Omron Sysmac Studio project Battery_System_Before_Test (Sysmac Studio 1.53.0.9, StandardProject)

# Controller new_Controller_0: NX102-1020 version 1.33
Units and slaves: 노드1 : NX-ECC203 (E005); 유니트 1 : NX-ID6142-6 (N8); 유니트 2 : NX-OD6121-6 (N9); 유니트 1 : NX-PF0730 (N1); 유니트 2 : NX-ILM400 (N2); 유니트 4 : NX-SID800 (N10); 유니트 5 : NX-SOD400 (N11)
Task PrimaryTask (priority 4, period or condition 2000): Program0, SlotTableProc

TYPE Slot_info : STRUCT
    SOC : UINT;  (* 배터리 잔량 % *)
    Status : INT;  (* 0 = 비어 있음 / 1 = 충전 중 / 2 = 불량 *)
    IO : WORD;  (* 로봇 신호 *)
END_STRUCT END_TYPE
TYPE U_IO16 : UNION
    W : WORD;
    B : ARRAY[0..15] OF BOOL;
END_UNION END_TYPE
TYPE S_RobotIO : STRUCT
    IO : U_IO16;
END_STRUCT END_TYPE

VAR_GLOBAL RETAIN
    Slot_No : ARRAY[1..6] OF Slot_Info := [(SOC := 16#0, Status := 1, IO := 16#01), (SOC := 16#0, Status := 1, IO := 16#02), (SOC := 16#0, Status := 1, IO := 16#04), (SOC := 16#0, Status := 1, IO := 16#08), (SOC := 16#0, Status := 1, IO := 16#10), (SOC := 16#0, Status := 1, IO := 16#20)];
END_VAR
VAR_GLOBAL
    Vision_Trigger : BOOL;  (* at ECAT://node#4/Line0 Trigger *)
    Vision_BC_Data : DINT;  (* at ECAT://node#4/Line0 DINT Result Data 0 *)
    Vision_Counter : DINT;  (* at ECAT://node#4/Line0 DINT Result Data 1 *)
    Robot_Send : S_RobotIO;
    Robot_Recv : S_RobotIO;
    MFC_HR : ARRAY[0..99] OF WORD;  (* PLC > MFC *)
    Arduino_HR : ARRAY[0..99] OF WORD;  (* Arduino > PLC *)
    Robot_In : ARRAY[0..237] OF WORD;  (* Robot > PLC; network input *)
    Robot_Out : ARRAY[0..105] OF WORD;  (* PLC > Robot; network output *)
    E_RST : BOOL;  (* Error Reset *)
    H_Rent_PB : BOOL;
    H_Card_Can_PB : BOOL;
    H_LowBatt_OK_PB : BOOL;
    H_LowBatt_Can_PB : BOOL;
    STP_D_SS : BOOL;  (* at ECAT://node#[1,1]/Input Bit 32 bits/Input Bit 16 *)
    STP_U_SS : BOOL;  (* at ECAT://node#[1,1]/Input Bit 32 bits/Input Bit 15 *)
    Detect_Home_SS : BOOL;  (* at ECAT://node#[1,1]/Input Bit 32 bits/Input Bit 22 *)
    Detect_STP_SS : BOOL;  (* at ECAT://node#[1,1]/Input Bit 32 bits/Input Bit 21 *)
    H_Vis_Rty_PB : BOOL;
    H_Vis_Home_PB : BOOL;
    H_Rtn_PB : BOOL;
    H_Rtn_Can_PB : BOOL;
    H_Refund_Can_PB : BOOL;
    H_Pop_Card : BOOL;
    H_pop_Wait_Rent : BOOL;
    H_Pop_LowBatt : BOOL;
    H_Pop_ContAdmin : BOOL;
    H_Pop_Rent_Done : BOOL;
    H_Pop_Place_Batt : BOOL;
    H_Pop_ReplBatt : BOOL;
    H_Pop_Refund : BOOL;
    H_Pop_RtnDone : BOOL;
    H_Pop_Equip_Running : BOOL;
    STP_SOL : BOOL;  (* at ECAT://node#[1,2]/Output Bit 32 bits/Output Bit 11 *)
    H_Scr_Main : BOOL;
    MotS_Status : WORD;  (* at ECAT://node#2/Status *)
    MotS : WORD;  (* at ECAT://node#2/Command *)
    MotM : WORD;  (* at ECAT://node#3/Command *)
    MotM_Status : WORD;  (* at ECAT://node#3/Status *)
    Batt_UseTime : ARRAY[1..6] OF TIME;
    Batt_Max_SOC : UINT;
    H_Pop_PayFail : BOOL;
    H_PayRty_PB : BOOL;
    H_PayFail_Home_PB : BOOL;
    Rtn_BC_IDX : DINT;
    Batt_Refund : LINT;
    H_Rst_PB : BOOL;
    H_Admin_PB : BOOL;
    H_Pop_Admin : BOOL;
    H_Admin_Home_PB : BOOL;
    RobotDone : BOOL;  (* 로봇 작업 완료 *)
    RobotMode : INT;  (* 1 : 반납 / 2 : 대여 *)
    RobotSlot : INT;  (* 로봇이 작업한 슬롯 번호 *)
    TestPctMode : BOOL;
    VisionBatteryID : WORD;  (* 바코드로 인식한 배터리 ID *)
    Batt_UseDisp : ARRAY[1..6] OF DINT;
    Batt_UseFee : LINT;
END_VAR

(* Program Program0: safety or other program stored in binary form, left out *)

PROGRAM Program0
VAR
    i : INT;
    Main_Process : FB_Batt_Process;
    MFC_ErrID : WORD;
    MFC_ReqCnt : UDINT;
    MFC : Connect;
    Arduino_Conn : BOOL;
    Arduino_ErrID : WORD;
    Arduino_ReqCnt : UDINT;
    Arduino : Connect;
    RPE : ResetPLCError;
    REE : ResetECError;
    RME : ResetMCError;
    Ard_PayOK : BOOL;
    Bot_Server_On : BOOL;
    First_Step : BOOL;
    T0 : TON;
    T1 : TON;
    C_Admin : CTU;
    T_Admin : TON;
END_VAR
VAR_EXTERNAL
    Slot_No : ARRAY[1..6] OF Slot_Info;
    Vision_BC_Data : DINT;
    MFC_HR : ARRAY[0..99] OF WORD;
    Arduino_HR : ARRAY[0..99] OF WORD;
    Robot_In : ARRAY[0..237] OF WORD;
    E_RST : BOOL;
    Vision_Counter : DINT;
    Robot_Recv : S_RobotIO;
    Robot_Send : S_RobotIO;
    Vision_Trigger : BOOL;
    H_Rent_PB : BOOL;
    H_Card_Can_PB : BOOL;
    H_LowBatt_OK_PB : BOOL;
    H_LowBatt_Can_PB : BOOL;
    STP_D_SS : BOOL;
    STP_U_SS : BOOL;
    Detect_Home_SS : BOOL;
    Detect_STP_SS : BOOL;
    H_Vis_Rty_PB : BOOL;
    H_Vis_Home_PB : BOOL;
    H_Rtn_PB : BOOL;
    H_Rtn_Can_PB : BOOL;
    H_Refund_Can_PB : BOOL;
    H_Pop_Card : BOOL;
    H_pop_Wait_Rent : BOOL;
    H_Pop_LowBatt : BOOL;
    H_Pop_ContAdmin : BOOL;
    H_Pop_Rent_Done : BOOL;
    H_Pop_Place_Batt : BOOL;
    H_Pop_ReplBatt : BOOL;
    H_Pop_Refund : BOOL;
    H_Pop_RtnDone : BOOL;
    H_Pop_Equip_Running : BOOL;
    STP_SOL : BOOL;
    H_Scr_Main : BOOL;
    MotM_Status : WORD;
    MotS_Status : WORD;
    MotM : WORD;
    MotS : WORD;
    Robot_Out : ARRAY[0..105] OF WORD;
    Batt_Max_SOC : UINT;
    H_Pop_PayFail : BOOL;
    H_PayRty_PB : BOOL;
    H_PayFail_Home_PB : BOOL;
    Rtn_BC_IDX : DINT;
    Batt_Refund : LINT;
    H_Rst_PB : BOOL;
    H_Admin_PB : BOOL;
    H_Pop_Admin : BOOL;
    H_Admin_Home_PB : BOOL;
    Batt_UseDisp : ARRAY[1..6] OF DINT;
    Batt_UseTime : ARRAY[1..6] OF TIME;
    Batt_UseFee : LINT;
END_VAR
VAR
    _e1 : R_TRIG;
    _e2 : R_TRIG;
END_VAR

(* Section Main_Program: ladder, written here as Structured Text *)

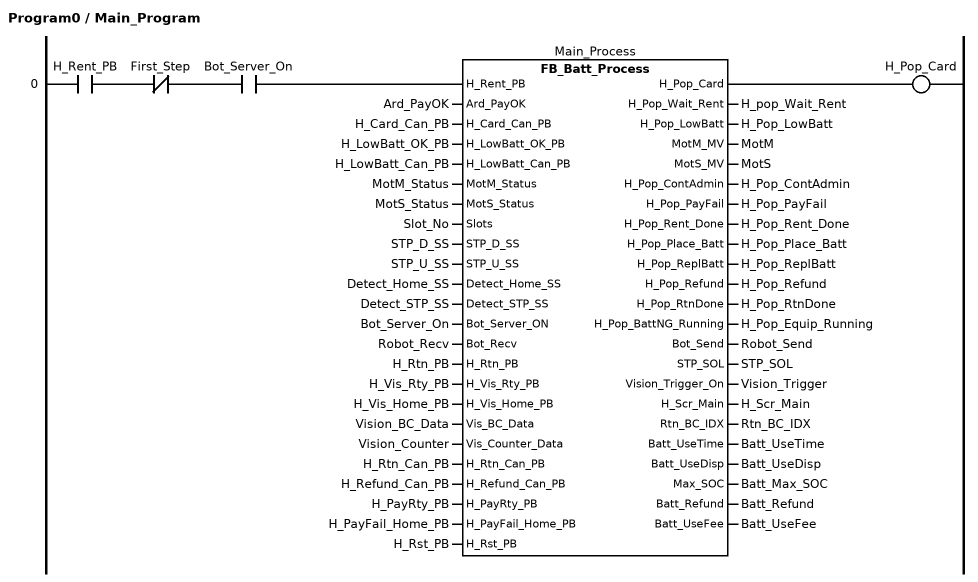
(* Rung 0 *)
Main_Process(H_Rent_PB := H_Rent_PB AND NOT First_Step AND Bot_Server_On, Ard_PayOK := Ard_PayOK, H_Card_Can_PB := H_Card_Can_PB, H_LowBatt_OK_PB := H_LowBatt_OK_PB, H_LowBatt_Can_PB := H_LowBatt_Can_PB, MotM_Status := MotM_Status, MotS_Status := MotS_Status, Slots := Slot_No, STP_D_SS := STP_D_SS, STP_U_SS := STP_U_SS, Detect_Home_SS := Detect_Home_SS, Detect_STP_SS := Detect_STP_SS, Bot_Server_ON := Bot_Server_On, Bot_Recv := Robot_Recv, H_Rtn_PB := H_Rtn_PB, H_Vis_Rty_PB := H_Vis_Rty_PB, H_Vis_Home_PB := H_Vis_Home_PB, Vis_BC_Data := Vision_BC_Data, Vis_Counter_Data := Vision_Counter, H_Rtn_Can_PB := H_Rtn_Can_PB, H_Refund_Can_PB := H_Refund_Can_PB, H_PayRty_PB := H_PayRty_PB, H_PayFail_Home_PB := H_PayFail_Home_PB, H_Rst_PB := H_Rst_PB, H_Pop_Wait_Rent => H_pop_Wait_Rent, H_Pop_LowBatt => H_Pop_LowBatt, MotM_MV => MotM, MotS_MV => MotS, H_Pop_ContAdmin => H_Pop_ContAdmin, H_Pop_PayFail => H_Pop_PayFail, H_Pop_Rent_Done => H_Pop_Rent_Done, H_Pop_Place_Batt => H_Pop_Place_Batt, H_Pop_ReplBatt => H_Pop_ReplBatt, H_Pop_Refund => H_Pop_Refund, H_Pop_RtnDone => H_Pop_RtnDone, H_Pop_BattNG_Running => H_Pop_Equip_Running, Bot_Send => Robot_Send, STP_SOL => STP_SOL, Vision_Trigger_On => Vision_Trigger, H_Scr_Main => H_Scr_Main, Rtn_BC_IDX => Rtn_BC_IDX, Batt_UseTime => Batt_UseTime, Batt_UseDisp => Batt_UseDisp, Max_SOC => Batt_Max_SOC, Batt_Refund => Batt_Refund, Batt_UseFee => Batt_UseFee);
H_Pop_Card := Main_Process.H_Pop_Card;

(* Section Sec_SOC_Copy: ladder, written here as Structured Text *)

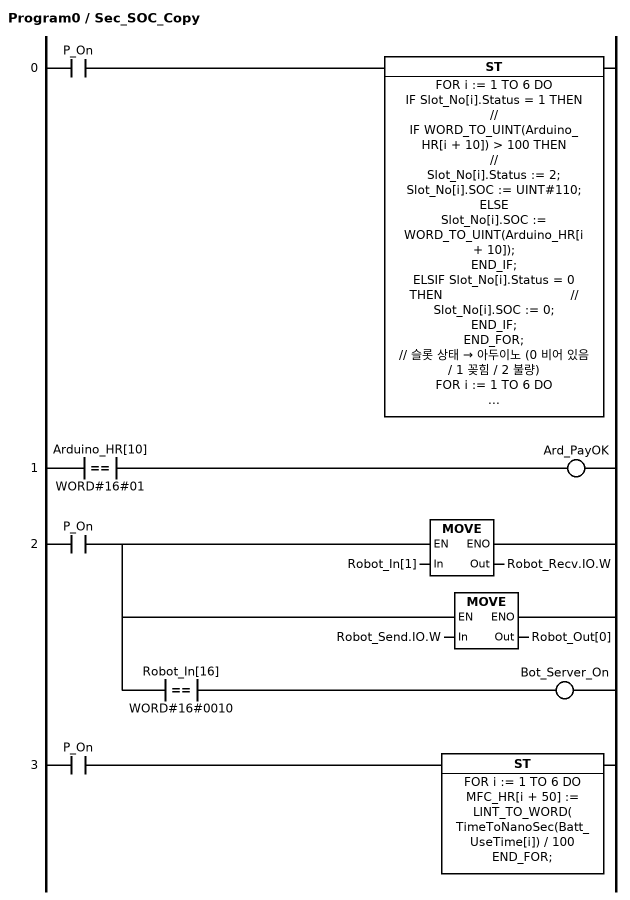
(* Rung 0 *)
IF P_On THEN
    FOR i := 1 TO 6 DO
        IF Slot_No[i].Status = 1 THEN                                   // 배터리가 꽂혀 있는 슬롯만 판단
            IF WORD_TO_UINT(Arduino_HR[i + 10]) > 100 THEN              // 아두이노 불량(110)
                Slot_No[i].Status := 2;
                Slot_No[i].SOC := UINT#110;
            ELSE
                Slot_No[i].SOC := WORD_TO_UINT(Arduino_HR[i + 10]);
            END_IF;
        ELSIF Slot_No[i].Status = 0 THEN                                // 빈 슬롯은 아두이노 값을 무시
            Slot_No[i].SOC := 0;
        END_IF;
    END_FOR;
    
    // 슬롯 상태 → 아두이노 (0 비어 있음 / 1 꽂힘 / 2 불량)
    FOR i := 1 TO 6 DO
        Arduino_HR[16 + i] := INT_TO_WORD(Slot_No[i].Status);
    END_FOR;
END_IF;
(* Rung 1 *)
Ard_PayOK := Arduino_HR[10] = WORD#16#01;
(* Rung 2 *)
IF P_On THEN
    Robot_Recv.IO.W := Robot_In[1];
    Robot_Out[0] := Robot_Send.IO.W;
END_IF;
Bot_Server_On := P_On AND (Robot_In[16] = WORD#16#0010);
(* Rung 3 *)
IF P_On THEN
    FOR i := 1 TO 6 DO
    	MFC_HR[i + 50] := LINT_TO_WORD( TimeToNanoSec(Batt_UseTime[i]) / 1000000000 );
    END_FOR;
END_IF;

(* Section Network: ladder, written here as Structured Text *)

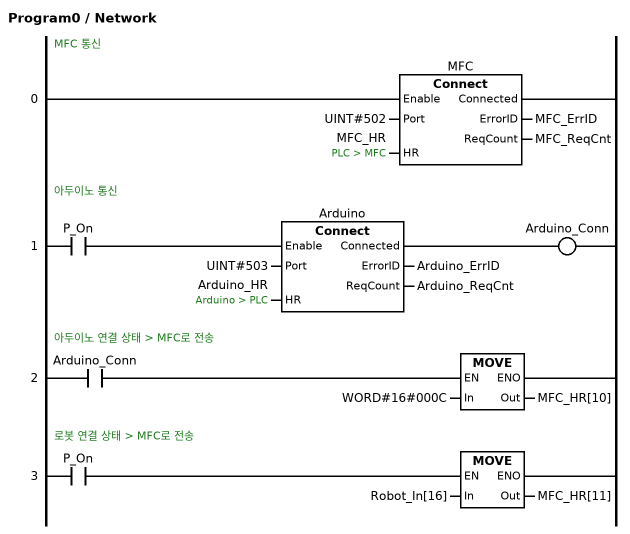
(* Rung 0: MFC 통신 *)
MFC(Enable := TRUE, Port := UINT#502, HR := MFC_HR, ErrorID => MFC_ErrID, ReqCount => MFC_ReqCnt);
(* Rung 1: 아두이노 통신 *)
Arduino(Enable := P_On, Port := UINT#503, HR := Arduino_HR, ErrorID => Arduino_ErrID, ReqCount => Arduino_ReqCnt);
Arduino_Conn := Arduino.Connected;
(* Rung 2: 아두이노 연결 상태 > MFC로 전송 *)
IF Arduino_Conn THEN MFC_HR[10] := WORD#16#000C; END_IF;
(* Rung 3: 로봇 연결 상태 > MFC로 전송 *)
IF P_On THEN MFC_HR[11] := Robot_In[16]; END_IF;

(* Section PLC_Error: ladder, written here as Structured Text *)

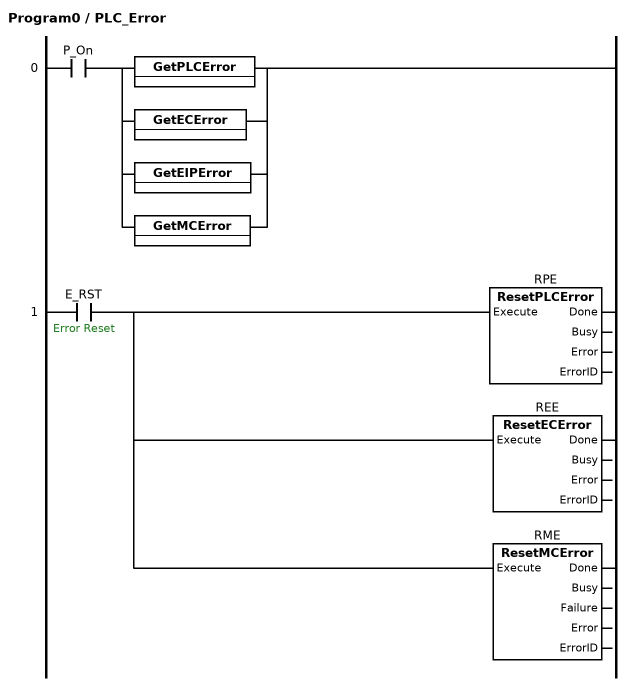
(* Rung 0 *)
(* drawn but driving nothing: P_On *)
(* Rung 1 *)
RPE(Execute := E_RST);
REE(Execute := E_RST);
RME(Execute := E_RST);

(* Section First_Scan: ladder, written here as Structured Text *)

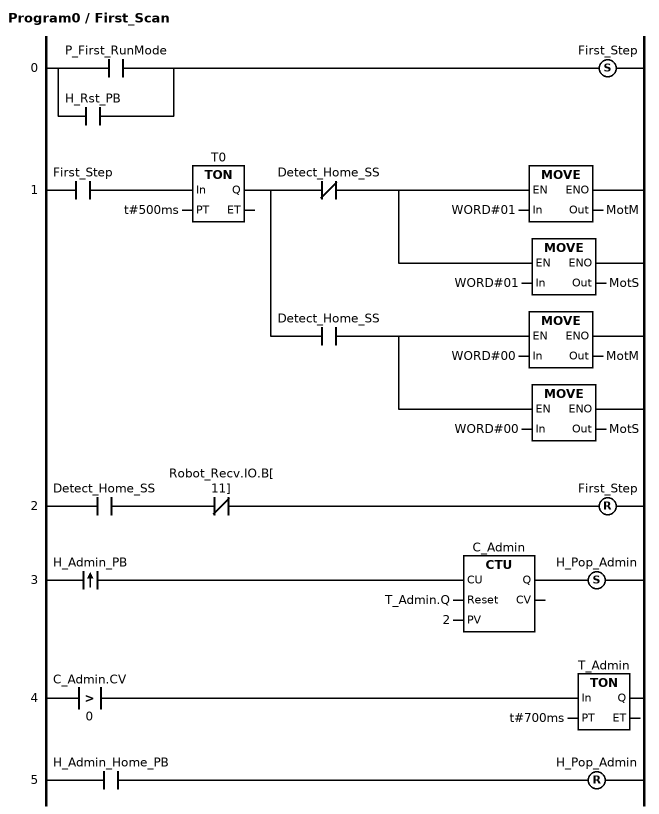
(* Rung 0 *)
IF P_First_RunMode OR H_Rst_PB THEN First_Step := TRUE; END_IF;
(* Rung 1 *)
T0(In := First_Step, PT := t#500ms);
IF T0.Q AND NOT Detect_Home_SS THEN
    MotM := WORD#01;
    MotS := WORD#01;
END_IF;
IF T0.Q AND Detect_Home_SS THEN
    MotM := WORD#00;
    MotS := WORD#00;
END_IF;
(* Rung 2 *)
IF Detect_Home_SS AND NOT Robot_Recv.IO.B[11] THEN First_Step := FALSE; END_IF;
(* Rung 3 *)
_e1(CLK := H_Admin_PB);
_e2(CLK := _e1.Q);
C_Admin(CU := _e2.Q, Reset := T_Admin.Q, PV := 2);
IF C_Admin.Q THEN H_Pop_Admin := TRUE; END_IF;
(* Rung 4 *)
T_Admin(In := C_Admin.CV > 0, PT := t#700ms);
(* Rung 5 *)
IF H_Admin_Home_PB THEN H_Pop_Admin := FALSE; END_IF;
END_PROGRAM

PROGRAM SlotTableProc
VAR
    i : INT;
    RentTrig : R_TRIG;
    ReturnTrig : R_TRIG;
    GripOnTrig : R_TRIG;
    GripOffTrig : F_TRIG;
    RobotKind : INT;
    RobotStep : INT;
    TestRobotMode : BOOL;
    TestRobotKind : INT;
    TestRobotStep : INT;
    GripState : BOOL;
    ErrTrig : R_TRIG;
    SlotNow : INT;
    SlotBitCnt : INT;
    ReturnCnt : UINT;
    RentCnt : UINT;
    RobotDO : WORD;
    DoRent : BOOL;
    DoReturn : BOOL;
    DoErr : BOOL;
    DoGripOn : BOOL;
    DoGripOff : BOOL;
    DoMove : BOOL;
    DoTask : BOOL;
    MoveTrig : R_TRIG;
    TaskEndTrig : F_TRIG;
    InitTrig : R_TRIG;
    InitMapping : BOOL;
END_VAR
VAR RETAIN
    SlotBatID : ARRAY[1..6] OF DINT := [1, 2, 3, 4, 5, 6];
END_VAR
VAR
    ReturnBatID : DINT;
END_VAR
VAR_EXTERNAL
    RobotDone : BOOL;
    RobotMode : INT;
    RobotSlot : INT;
    Vision_BC_Data : DINT;
    MFC_HR : ARRAY[0..99] OF WORD;
    Slot_No : ARRAY[1..6] OF Slot_Info;
    Arduino_HR : ARRAY[0..99] OF WORD;
    TestPctMode : BOOL;
    Robot_In : ARRAY[0..237] OF WORD;
    Robot_Out : ARRAY[0..105] OF WORD;
END_VAR
// ───── 0. 시연 시작 : 슬롯 n = 배터리 n 으로 초기 등록 (InitMapping 을 켤 때만) ─────
InitTrig(Clk := InitMapping);
IF InitTrig.Q THEN
    FOR i := 1 TO 6 DO
        SlotBatID[i] := INT_TO_DINT(i);      // 슬롯 1 = 배터리 1 ...
        Slot_No[i].Status := 1;              // 전부 꽂혀 있는 상태로
    END_FOR;
    MFC_HR[46] := WORD#0;                    // 마지막 대여 배터리 ID 지움
END_IF;

// ───── 1. 로봇 DO (Robot_In[1]) → 작업 종류 / 슬롯 / 단계 ─────
RobotDO := Robot_In[1];

DoRent     := (RobotDO AND WORD#16#0040) <> WORD#0;   // DO7  대여
DoReturn   := (RobotDO AND WORD#16#0080) <> WORD#0;   // DO8  반납
DoErr      := (RobotDO AND WORD#16#0100) <> WORD#0;   // DO9  고장 회수
DoMove     := (RobotDO AND WORD#16#0400) <> WORD#0;   // DO11 이동 중 (집으러 / 놓으러)
DoGripOff  := (RobotDO AND WORD#16#4000) <> WORD#0;   // DO15 그리퍼 열기
DoGripOn   := (RobotDO AND WORD#16#8000) <> WORD#0;   // DO16 그리퍼 잡기
DoTask     := DoRent OR DoReturn OR DoErr;            // 작업 신호 중 하나라도 켜짐

RentTrig(Clk := DoRent);
ReturnTrig(Clk := DoReturn);
ErrTrig(Clk := DoErr);
MoveTrig(Clk := DoMove);
TaskEndTrig(Clk := DoTask);                           // F_TRIG : 로봇이 DO7/8/9 를 끄는 순간
 
// DO1~6 → 슬롯 번호 (딱 하나만 켜져 있을 때만 인정)
SlotNow := 0;
SlotBitCnt := 0;
FOR i := 0 TO 5 DO
    IF (RobotDO AND SHL(WORD#16#0001, INT_TO_UINT(i))) <> WORD#0 THEN
        SlotNow := i + 1;
        SlotBitCnt := SlotBitCnt + 1;
    END_IF;
END_FOR;
IF SlotBitCnt <> 1 THEN
    SlotNow := 0;
END_IF;

// 1단계 작업 접수 : DO7 / DO8 / DO9 켜짐
IF RentTrig.Q THEN
    RobotKind := 1; RobotMode := 2; RobotStep := 1; RobotSlot := 0;
END_IF;
IF ReturnTrig.Q THEN
    RobotKind := 2; RobotMode := 1; RobotStep := 1; RobotSlot := 0;
END_IF;
IF ErrTrig.Q THEN
    RobotKind := 3; RobotMode := 3; RobotStep := 1; RobotSlot := 0;
END_IF;

// 슬롯 번호 확정 (DO7/8/9와 DO1~6이 같은 스캔에 안 들어와도 잡히게)
IF (RobotKind >= 1) AND (RobotKind <= 3) AND (RobotSlot = 0) AND (SlotNow <> 0) THEN
    RobotSlot := SlotNow;
END_IF;

// 2단계 / 4단계 이동 : DO11 이 켜질 때마다
IF MoveTrig.Q THEN
    IF RobotStep = 1 THEN
        RobotStep := 2;                               // 첫 번째 이동 : 집으러 감
    ELSIF RobotStep = 3 THEN
        RobotStep := 4;                               // 두 번째 이동 : 놓으러 감
    END_IF;
END_IF;

// 3단계 파지 : DO16 잡기 켜짐 + DO15 열기 꺼짐
IF DoGripOn AND NOT DoGripOff AND (RobotStep = 2) THEN
    RobotStep := 3;
END_IF;

// 5단계 배출 / 삽입 : DO15 열기 켜짐 + DO16 잡기 꺼짐
IF DoGripOff AND NOT DoGripOn AND (RobotStep = 4) THEN
    RobotStep := 5;
END_IF;

// 6단계 완료 : 로봇이 DO7/8/9 를 끄는 순간
RobotDone := TaskEndTrig.Q AND (RobotStep = 5);
IF RobotDone THEN
    RobotStep := 6;
END_IF;

// ───── 2. 로봇 작업 완료 → 슬롯 상태 / 배터리 ID 갱신 ─────
IF RobotDone THEN
    IF (RobotSlot >= 1) AND (RobotSlot <= 6) THEN
        IF RobotMode = 1 THEN                                   // 반납 : 충전 중
			ReturnBatID := Vision_BC_Data;
            Slot_No[RobotSlot].Status := 1;
            SlotBatID[RobotSlot] := ReturnBatID;
            MFC_HR[14] := INT_TO_WORD(RobotSlot);               // 반납 슬롯
            ReturnCnt := ReturnCnt + 1;
            MFC_HR[15] := UINT_TO_WORD(ReturnCnt);              // 반납 횟수
        ELSIF RobotMode = 2 THEN                                // 대여 : 비움
            MFC_HR[46] := DINT_TO_WORD(SlotBatID[RobotSlot]);   // 지우기 전에 대여 배터리 ID 보관
            Slot_No[RobotSlot].SOC    := UINT#0;
            Slot_No[RobotSlot].Status := 0;
            SlotBatID[RobotSlot] := DINT#0;
            MFC_HR[12] := INT_TO_WORD(RobotSlot);               // 대여 슬롯
            RentCnt := RentCnt + 1;
            MFC_HR[13] := UINT_TO_WORD(RentCnt);                // 대여 횟수
        ELSIF RobotMode = 3 THEN                                // 고장 회수 : 비움
            Slot_No[RobotSlot].SOC    := UINT#0;
            Slot_No[RobotSlot].Status := 0;
            SlotBatID[RobotSlot] := DINT#0;
        END_IF;
    END_IF;
END_IF;

// (아두이노 잔량 → Slot_No[i].SOC 는 기존 Rung 0 에서 처리하므로 여기서 뺌)

// ───── 3. 슬롯 테이블 → MFC_HR[17]~[37] ─────
FOR i := 0 TO 6 DO
    MFC_HR[17 + i * 3] := INT_TO_WORD(Slot_No[i].Status);
    MFC_HR[18 + i * 3] := UINT_TO_WORD(Slot_No[i].SOC);     // SOC가 UINT라 WORD로 변환
    MFC_HR[19 + i * 3] := Slot_No[i].IO;
END_FOR;

// ───── 4. 로봇 작업 상태 → MFC_HR[38]~[39] ─────
MFC_HR[38] := INT_TO_WORD(RobotKind);       // 0 대기 / 1 대여 / 2 반납 / 3 고장 회수
MFC_HR[39] := INT_TO_WORD(RobotStep);       // 1 접수 / 2 이동 / 3 파지 / 4 이동 / 5 배출·삽입 / 6 완료

// ───── 5. 슬롯별 배터리 ID → MFC_HR[40]~[45] ─────
FOR i := 1 TO 6 DO
    MFC_HR[39 + i] := DINT_TO_WORD(SlotBatID[i]);
END_FOR;
END_PROGRAM

FUNCTION_BLOCK Hmi_Rent
VAR
    data : INT;
    W_RecMax_Pos : ARRAY[0..5] OF UINT;
    T0 : TON;
    T1 : TON;
END_VAR
VAR_INPUT
    Hmi_Start : BOOL;
END_VAR
VAR_OUTPUT
    H_Pop_Wait_Rent : BOOL;
END_VAR
VAR_INPUT
    Ard_PayOK : BOOL;
    Max_SOC : UINT;
END_VAR
VAR_OUTPUT
    H_Pop_Card : BOOL;
END_VAR
VAR_INPUT
    H_Card_Cancle_PB : BOOL;
END_VAR
VAR_OUTPUT
    H_Pop_LowBatt : BOOL;
END_VAR
VAR_INPUT
    H_LowBatt_OK_PB : BOOL;
    H_LowBatt_Can_PB : BOOL;
    H_PayRty_PB : BOOL;
    H_PayFail_Home_PB : BOOL;
    Cmd_Ack : BOOL;
END_VAR
VAR_OUTPUT
    H_Pop_PayFail : BOOL;
    Hmi_Busy : BOOL;
END_VAR
VAR_INPUT
    H_Rst_PB : BOOL;
END_VAR
VAR
    _e1 : R_TRIG;
    _p2 : BOOL;
    _p3 : BOOL;
    _p4 : BOOL;
    _p5 : BOOL;
END_VAR
(* ladder, written here as Structured Text *)

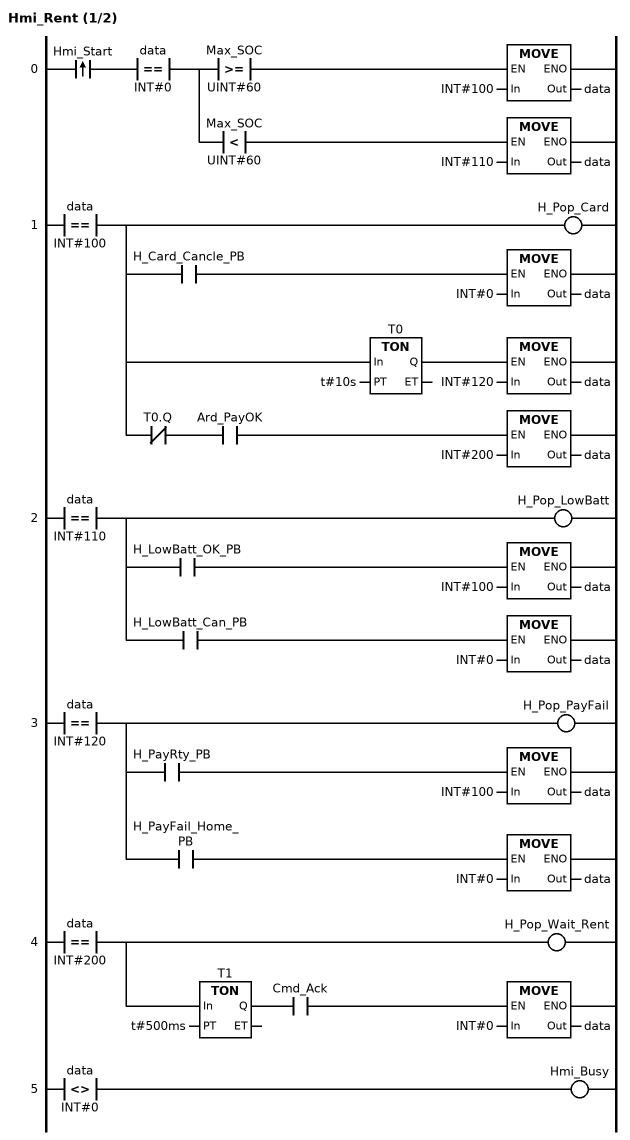
(* Rung 0 *)
_e1(CLK := Hmi_Start);
_p2 := _e1.Q AND (data = INT#0);
IF _e1.Q AND (data = INT#0) AND (Max_SOC >= UINT#60) THEN data := INT#100; END_IF;
IF _p2 AND (Max_SOC < UINT#60) THEN data := INT#110; END_IF;
(* Rung 1 *)
H_Pop_Card := data = INT#100;
_p3 := data = INT#100;
IF (data = INT#100) AND H_Card_Cancle_PB THEN data := INT#0; END_IF;
T0(In := _p3, PT := t#10s);
IF T0.Q THEN data := INT#120; END_IF;
IF _p3 AND NOT T0.Q AND Ard_PayOK THEN data := INT#200; END_IF;
(* Rung 2 *)
H_Pop_LowBatt := data = INT#110;
_p4 := data = INT#110;
IF (data = INT#110) AND H_LowBatt_OK_PB THEN data := INT#100; END_IF;
IF _p4 AND H_LowBatt_Can_PB THEN data := INT#0; END_IF;
(* Rung 3 *)
H_Pop_PayFail := data = INT#120;
_p5 := data = INT#120;
IF (data = INT#120) AND H_PayRty_PB THEN data := INT#100; END_IF;
IF _p5 AND H_PayFail_Home_PB THEN data := INT#0; END_IF;
(* Rung 4 *)
H_Pop_Wait_Rent := data = INT#200;
T1(In := data = INT#200, PT := t#500ms);
IF T1.Q AND Cmd_Ack THEN data := INT#0; END_IF;
(* Rung 5 *)
Hmi_Busy := data <> INT#0;

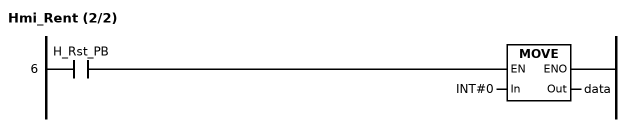
(* Rung 6 *)
IF H_Rst_PB THEN data := INT#0; END_IF;
END_FUNCTION_BLOCK

FUNCTION_BLOCK Robot_Move
VAR
    Cmd_Base : WORD;
    data : INT;
END_VAR
VAR_INPUT
    Bot_Start : BOOL;
END_VAR
VAR_OUTPUT
    Bot_Done : BOOL;
END_VAR
VAR_INPUT
    Bot_Server_On : BOOL;
    MPS_Ready : BOOL;
    Bot_Mode_IO : WORD;
    Bot_Recv : S_RobotIO;
    Target_Slot_NO : UINT;
END_VAR
VAR_OUTPUT
    Bot_Clear : BOOL;
    Bot_Send : S_RobotIO;
END_VAR
VAR_INPUT
    Cmd_Ack : BOOL;
END_VAR
VAR_IN_OUT
    Slots : ARRAY[1..6] OF Slot_info;
END_VAR
VAR_INPUT
    Slot_Status_data : INT;
END_VAR
VAR_OUTPUT
    Robot_Busy : BOOL;
END_VAR
VAR_INPUT
    H_Rst_PB : BOOL;
END_VAR
VAR
    _e1 : R_TRIG;
END_VAR
(* ladder, written here as Structured Text *)

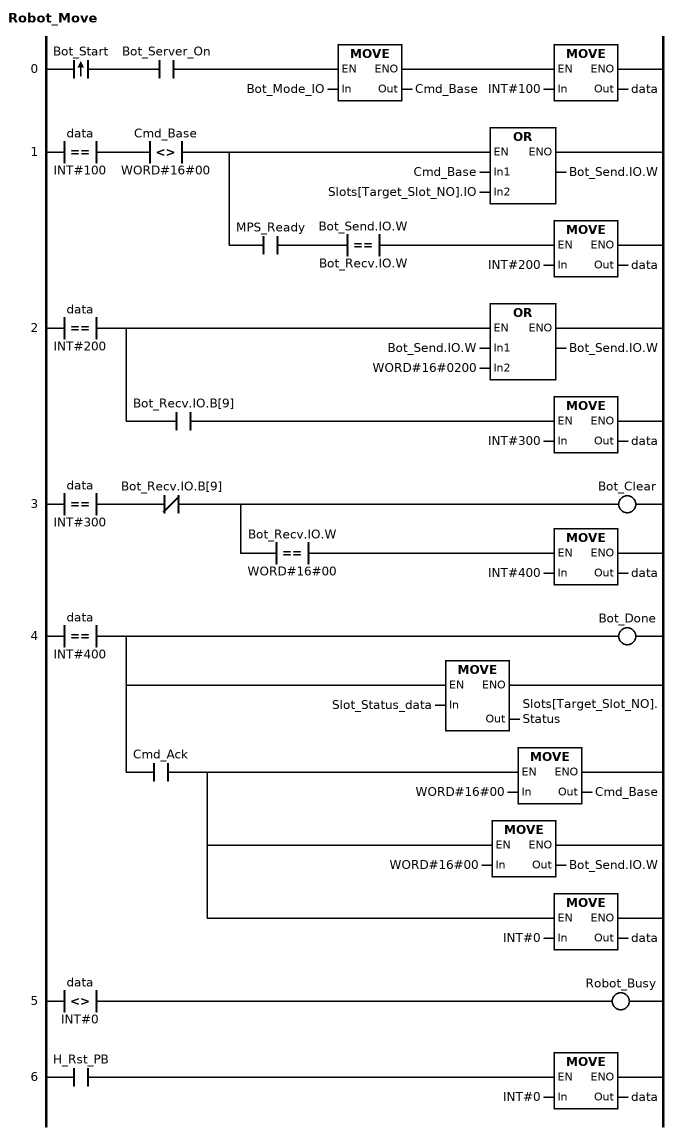
(* Rung 0 *)
_e1(CLK := Bot_Start);
IF _e1.Q AND Bot_Server_On THEN
    Cmd_Base := Bot_Mode_IO;
    data := INT#100;
END_IF;
(* Rung 1 *)
IF (data = INT#100) AND (Cmd_Base <> WORD#16#00) THEN
    Bot_Send.IO.W := Cmd_Base OR Slots[Target_Slot_NO].IO;
END_IF;
IF (data = INT#100) AND (Cmd_Base <> WORD#16#00) AND MPS_Ready AND (Bot_Send.IO.W = Bot_Recv.IO.W) THEN
    data := INT#200;
END_IF;
(* Rung 2 *)
IF data = INT#200 THEN Bot_Send.IO.W := Bot_Send.IO.W OR WORD#16#0200; END_IF;
IF (data = INT#200) AND Bot_Recv.IO.B[9] THEN data := INT#300; END_IF;
(* Rung 3 *)
Bot_Clear := (data = INT#300) AND NOT Bot_Recv.IO.B[9];
IF (data = INT#300) AND NOT Bot_Recv.IO.B[9] AND (Bot_Recv.IO.W = WORD#16#00) THEN
    data := INT#400;
END_IF;
(* Rung 4 *)
Bot_Done := data = INT#400;
IF data = INT#400 THEN Slots[Target_Slot_NO].Status := Slot_Status_data; END_IF;
IF (data = INT#400) AND Cmd_Ack THEN
    Cmd_Base := WORD#16#00;
    Bot_Send.IO.W := WORD#16#00;
    data := INT#0;
END_IF;
(* Rung 5 *)
Robot_Busy := data <> INT#0;
(* Rung 6 *)
IF H_Rst_PB THEN data := INT#0; END_IF;
END_FUNCTION_BLOCK

FUNCTION_BLOCK MPS
VAR
    data : INT;
END_VAR
VAR_INPUT
    MPS_Start : BOOL;
END_VAR
VAR_OUTPUT
    MPS_Done : BOOL;
END_VAR
VAR_INPUT
    MotM_Status : WORD;
    MotS_Status : WORD;
END_VAR
VAR_OUTPUT
    Motor_Run : BOOL;
    Sub_Motor_Run : BOOL;
END_VAR
VAR_INPUT
    STP_Start_SS : BOOL;
    STP_End_SS : BOOL;
END_VAR
VAR_OUTPUT
    STP_Sol : BOOL;
END_VAR
VAR_INPUT
    Detect_Start_SS : BOOL;
    Detect_End_SS : BOOL;
    Cmd_Ack : BOOL;
END_VAR
VAR_OUTPUT
    MPS_Busy : BOOL;
END_VAR
VAR_INPUT
    H_Rst_PB : BOOL;
END_VAR
VAR
    _e1 : R_TRIG;
    _p2 : BOOL;
END_VAR
(* ladder, written here as Structured Text *)

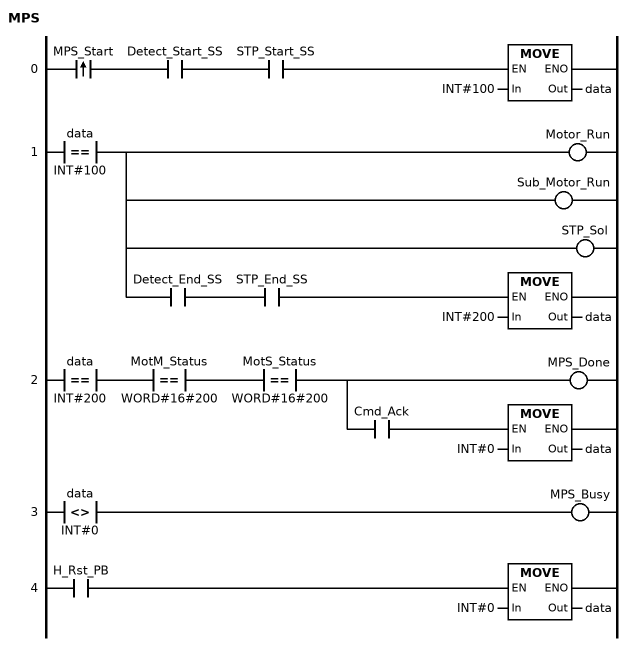
(* Rung 0 *)
_e1(CLK := MPS_Start);
IF _e1.Q AND Detect_Start_SS AND STP_Start_SS THEN data := INT#100; END_IF;
(* Rung 1 *)
Motor_Run := data = INT#100;
Sub_Motor_Run := data = INT#100;
STP_Sol := data = INT#100;
IF (data = INT#100) AND Detect_End_SS AND STP_End_SS THEN data := INT#200; END_IF;
(* Rung 2 *)
_p2 := (data = INT#200) AND (MotM_Status = WORD#16#200) AND (MotS_Status = WORD#16#200);
MPS_Done := _p2;
IF _p2 AND Cmd_Ack THEN data := INT#0; END_IF;
(* Rung 3 *)
MPS_Busy := data <> INT#0;
(* Rung 4 *)
IF H_Rst_PB THEN data := INT#0; END_IF;
END_FUNCTION_BLOCK

FUNCTION_BLOCK Rent
VAR
    Rent_Robot : Robot_Move;
    H_Rent : Hmi_Rent;
    Vision_Rent : Vision;
    T0 : TON;
    data : INT;
    MAX_Data : RecMax_Data;
    RecMax_Done : BOOL;
    Vision_Done : BOOL;
    Rent_Eq_Cycle : FB_Equipment_Cycle;
    Eq_Cycle_Done : BOOL;
    Max_Slot_No : UINT;
    Vis_Busy : BOOL;
    Equip_Busy : BOOL;
    Hmi_Busy : BOOL;
    T1 : TON;
END_VAR
VAR_INPUT
    Rent_Start : BOOL;
    Ard_PayOK : BOOL;
    H_Card_Can_PB : BOOL;
    H_LowBatt_OK_PB : BOOL;
    H_LowBatt_Can_PB : BOOL;
END_VAR
VAR_OUTPUT
    H_Pop_Card : BOOL;
    H_Pop_Wait_Rent : BOOL;
    H_Pop_LowBatt : BOOL;
END_VAR
VAR_INPUT
    MotM_Status : WORD;
    MotS_Status : WORD;
END_VAR
VAR_OUTPUT
    MotM_CCW : BOOL;
    MotS_CW : BOOL;
    MotS_CCW : BOOL;
    MotM_CW : BOOL;
END_VAR
VAR_IN_OUT
    Slots : ARRAY[1..6] OF Slot_info;
END_VAR
VAR_OUTPUT
    Bot_Send : S_RobotIO;
END_VAR
VAR_INPUT
    STP_D_SS : BOOL;
    STP_U_SS : BOOL;
END_VAR
VAR_OUTPUT
    STP_SOL : BOOL;
END_VAR
VAR_INPUT
    Detect_Home_SS : BOOL;
    Detect_STP_SS : BOOL;
    Vision_BC_Data : DINT;
    Vision_Counter_Data : DINT;
END_VAR
VAR_OUTPUT
    Vision_On : BOOL;
    H_Pop_ContAdmin : BOOL;
END_VAR
VAR_INPUT
    H_Vision_Rty_PB : BOOL;
    H_Vision_Home_PB : BOOL;
    H_PayRty_PB : BOOL;
END_VAR
VAR_OUTPUT
    H_Pop_Rent_Done : BOOL;
END_VAR
VAR_INPUT
    H_PayFail_Home_PB : BOOL;
END_VAR
VAR_OUTPUT
    H_Pop_PayFail : BOOL;
    BC_IDX_NO : DINT;
END_VAR
VAR_INPUT
    Bot_Server_On : BOOL;
    Bot_Recv : S_RobotIO;
END_VAR
VAR_OUTPUT
    Rent_Busy : BOOL;
    H_Scr_Main : BOOL;
    Batt_UseStart : BOOL;
    Max_SOC : UINT;
END_VAR
VAR_INPUT
    H_Rst_PB : BOOL;
END_VAR
(* ladder, written here as Structured Text *)

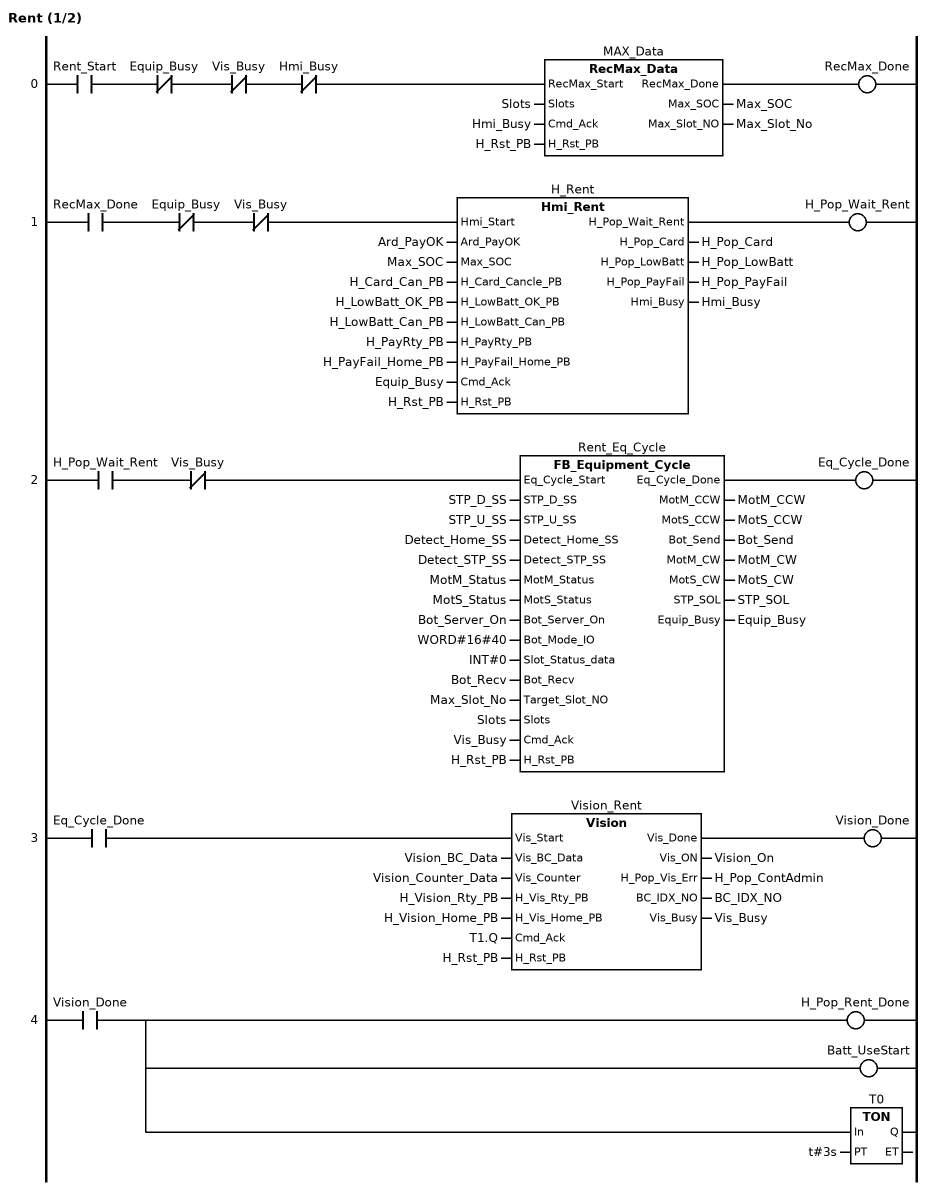
(* Rung 0 *)
MAX_Data(RecMax_Start := Rent_Start AND NOT Equip_Busy AND NOT Vis_Busy AND NOT Hmi_Busy, Slots := Slots, Cmd_Ack := Hmi_Busy, H_Rst_PB := H_Rst_PB, Max_SOC => Max_SOC, Max_Slot_NO => Max_Slot_No);
RecMax_Done := MAX_Data.RecMax_Done;
(* Rung 1 *)
H_Rent(Hmi_Start := RecMax_Done AND NOT Equip_Busy AND NOT Vis_Busy, Ard_PayOK := Ard_PayOK, Max_SOC := Max_SOC, H_Card_Cancle_PB := H_Card_Can_PB, H_LowBatt_OK_PB := H_LowBatt_OK_PB, H_LowBatt_Can_PB := H_LowBatt_Can_PB, H_PayRty_PB := H_PayRty_PB, H_PayFail_Home_PB := H_PayFail_Home_PB, Cmd_Ack := Equip_Busy, H_Rst_PB := H_Rst_PB, H_Pop_Card => H_Pop_Card, H_Pop_LowBatt => H_Pop_LowBatt, H_Pop_PayFail => H_Pop_PayFail, Hmi_Busy => Hmi_Busy);
H_Pop_Wait_Rent := H_Rent.H_Pop_Wait_Rent;
(* Rung 2 *)
Rent_Eq_Cycle(Eq_Cycle_Start := H_Pop_Wait_Rent AND NOT Vis_Busy, STP_D_SS := STP_D_SS, STP_U_SS := STP_U_SS, Detect_Home_SS := Detect_Home_SS, Detect_STP_SS := Detect_STP_SS, MotM_Status := MotM_Status, MotS_Status := MotS_Status, Bot_Server_On := Bot_Server_On, Bot_Mode_IO := WORD#16#40, Slot_Status_data := INT#0, Bot_Recv := Bot_Recv, Target_Slot_NO := Max_Slot_No, Slots := Slots, Cmd_Ack := Vis_Busy, H_Rst_PB := H_Rst_PB, MotM_CCW => MotM_CCW, MotS_CCW => MotS_CCW, Bot_Send => Bot_Send, MotM_CW => MotM_CW, MotS_CW => MotS_CW, STP_SOL => STP_SOL, Equip_Busy => Equip_Busy);
Eq_Cycle_Done := Rent_Eq_Cycle.Eq_Cycle_Done;
(* Rung 3 *)
Vision_Rent(Vis_Start := Eq_Cycle_Done, Vis_BC_Data := Vision_BC_Data, Vis_Counter := Vision_Counter_Data, H_Vis_Rty_PB := H_Vision_Rty_PB, H_Vis_Home_PB := H_Vision_Home_PB, Cmd_Ack := T1.Q, H_Rst_PB := H_Rst_PB, Vis_ON => Vision_On, H_Pop_Vis_Err => H_Pop_ContAdmin, BC_IDX_NO => BC_IDX_NO, Vis_Busy => Vis_Busy);
Vision_Done := Vision_Rent.Vis_Done;
(* Rung 4 *)
H_Pop_Rent_Done := Vision_Done;
Batt_UseStart := Vision_Done;
T0(In := Vision_Done, PT := t#3s);

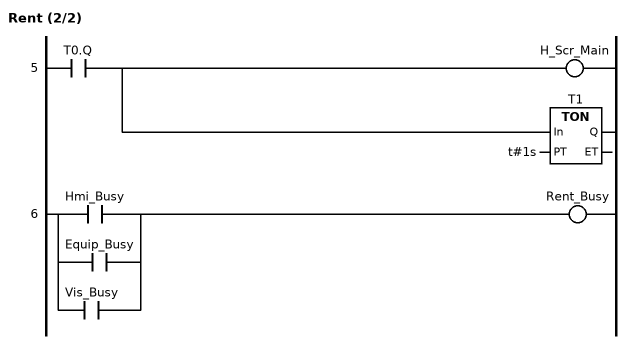
(* Rung 5 *)
H_Scr_Main := T0.Q;
T1(In := T0.Q, PT := t#1s);
(* Rung 6 *)
Rent_Busy := Hmi_Busy OR Equip_Busy OR Vis_Busy;
END_FUNCTION_BLOCK

FUNCTION_BLOCK Vision
VAR
    data : INT;
    T0 : TON;
    Old_Vis_Counter : DINT;
    C0 : CTU;
    C0_Rst : BOOL;
    T1 : TON;
END_VAR
VAR_INPUT
    Vis_Start : BOOL;
END_VAR
VAR_OUTPUT
    Vis_Done : BOOL;
    Vis_ON : BOOL;
END_VAR
VAR_INPUT
    Vis_BC_Data : DINT;
    Vis_Counter : DINT;
END_VAR
VAR_OUTPUT
    H_Pop_Vis_Err : BOOL;
END_VAR
VAR_INPUT
    H_Vis_Rty_PB : BOOL;
    H_Vis_Home_PB : BOOL;
END_VAR
VAR_OUTPUT
    BC_IDX_NO : DINT;
END_VAR
VAR_INPUT
    Cmd_Ack : BOOL;
END_VAR
VAR_OUTPUT
    Vis_Busy : BOOL;
END_VAR
VAR_INPUT
    H_Rst_PB : BOOL;
END_VAR
VAR
    _e1 : R_TRIG;
    _p2 : BOOL;
    _e3 : R_TRIG;
    _p4 : BOOL;
    _p5 : BOOL;
END_VAR
(* ladder, written here as Structured Text *)

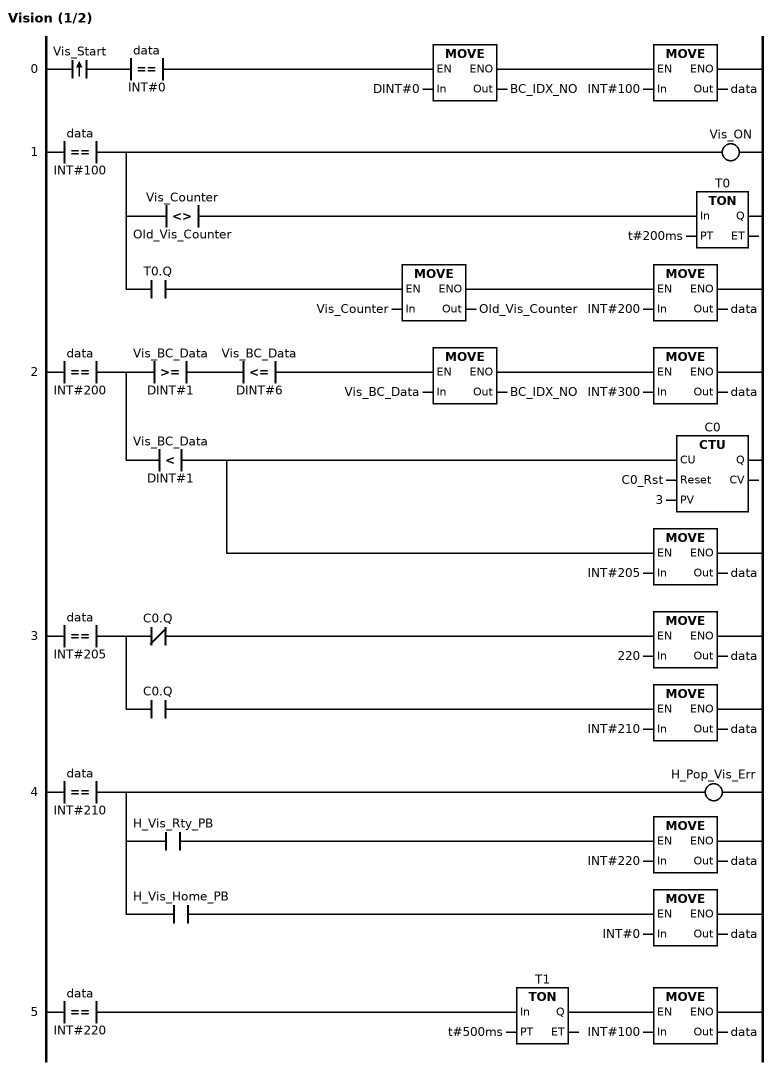
(* Rung 0 *)
_e1(CLK := Vis_Start);
IF _e1.Q AND (data = INT#0) THEN
    BC_IDX_NO := DINT#0;
    data := INT#100;
END_IF;
(* Rung 1 *)
Vis_ON := data = INT#100;
T0(In := (data = INT#100) AND (Vis_Counter <> Old_Vis_Counter), PT := t#200ms);
IF (data = INT#100) AND T0.Q THEN
    Old_Vis_Counter := Vis_Counter;
    data := INT#200;
END_IF;
(* Rung 2 *)
IF (data = INT#200) AND (Vis_BC_Data >= DINT#1) AND (Vis_BC_Data <= DINT#6) THEN
    BC_IDX_NO := Vis_BC_Data;
END_IF;
_p2 := data = INT#200;
IF (data = INT#200) AND (Vis_BC_Data >= DINT#1) AND (Vis_BC_Data <= DINT#6) THEN data := INT#300; END_IF;
_e3(CLK := _p2 AND (Vis_BC_Data < DINT#1));
C0(CU := _e3.Q, Reset := C0_Rst, PV := 3);
IF _p2 AND (Vis_BC_Data < DINT#1) THEN data := INT#205; END_IF;
(* Rung 3 *)
_p4 := data = INT#205;
IF (data = INT#205) AND NOT C0.Q THEN data := 220; END_IF;
IF _p4 AND C0.Q THEN data := INT#210; END_IF;
(* Rung 4 *)
H_Pop_Vis_Err := data = INT#210;
_p5 := data = INT#210;
IF (data = INT#210) AND H_Vis_Rty_PB THEN data := INT#220; END_IF;
IF _p5 AND H_Vis_Home_PB THEN data := INT#0; END_IF;
(* Rung 5 *)
T1(In := data = INT#220, PT := t#500ms);
IF T1.Q THEN data := INT#100; END_IF;

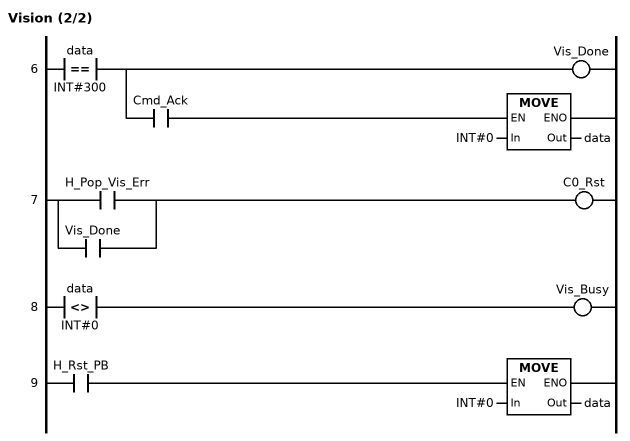
(* Rung 6 *)
Vis_Done := data = INT#300;
IF (data = INT#300) AND Cmd_Ack THEN data := INT#0; END_IF;
(* Rung 7 *)
C0_Rst := H_Pop_Vis_Err OR Vis_Done;
(* Rung 8 *)
Vis_Busy := data <> INT#0;
(* Rung 9 *)
IF H_Rst_PB THEN data := INT#0; END_IF;
END_FUNCTION_BLOCK

FUNCTION_BLOCK Rtn
VAR
    Empty_Slot_Data : RecSearch_Data;
    RecSrch_Done : BOOL;
    Empty_Slot_NO : UINT;
    H_Rtn : Hmi_Rtn;
    Rtn_Eq_Cycle : FB_Equipment_Cycle;
    Eq_Cycle_Done : BOOL;
    T0 : TON;
    Hmi_Rtn_Busy : BOOL;
    Equip_Busy : BOOL;
    T1 : TON;
END_VAR
VAR_INPUT
    Rtn_Start : BOOL;
END_VAR
VAR_IN_OUT
    Slots : ARRAY[1..6] OF Slot_info;
END_VAR
VAR_INPUT
    H_Vis_Rty_PB : BOOL;
    H_Vis_Home_PB : BOOL;
    Vis_BC_Data : DINT;
    Vis_Counter : DINT;
    Ard_PayOK : BOOL;
END_VAR
VAR_OUTPUT
    H_Pop_PlaceBatt : BOOL;
    Vis_On : BOOL;
    H_Pop_ReplBatt : BOOL;
    BC_IDX_NO : DINT;
    H_Pop_Refund : BOOL;
    H_Pop_PayFail : BOOL;
    H_Pop_RtnDone : BOOL;
END_VAR
VAR_INPUT
    H_Rtn_Can_PB : BOOL;
    H_Refund_Can_PB : BOOL;
    H_PayFail_Home_PB : BOOL;
    H_PayRty_PB : BOOL;
    MotM_Status : WORD;
    MotS_Status : WORD;
END_VAR
VAR_OUTPUT
    MotM_CCW : BOOL;
    MotS_CCW : BOOL;
    MotM_CW : BOOL;
    MotS_CW : BOOL;
END_VAR
VAR_INPUT
    STP_D_SS : BOOL;
    STP_U_SS : BOOL;
    Detect_Home_SS : BOOL;
    Detect_STP_SS : BOOL;
    Bot_Server_On : BOOL;
    Bot_Recv : S_RobotIO;
END_VAR
VAR_OUTPUT
    Bot_Send : S_RobotIO;
    STP_SOL : BOOL;
    H_Scr_Main : BOOL;
    Rtn_Busy : BOOL;
    Batt_UseDone : BOOL;
    Rtn_Equip_Running : BOOL;
END_VAR
VAR_INPUT
    H_Rst_PB : BOOL;
END_VAR
VAR
    _p1 : BOOL;
END_VAR
(* ladder, written here as Structured Text *)

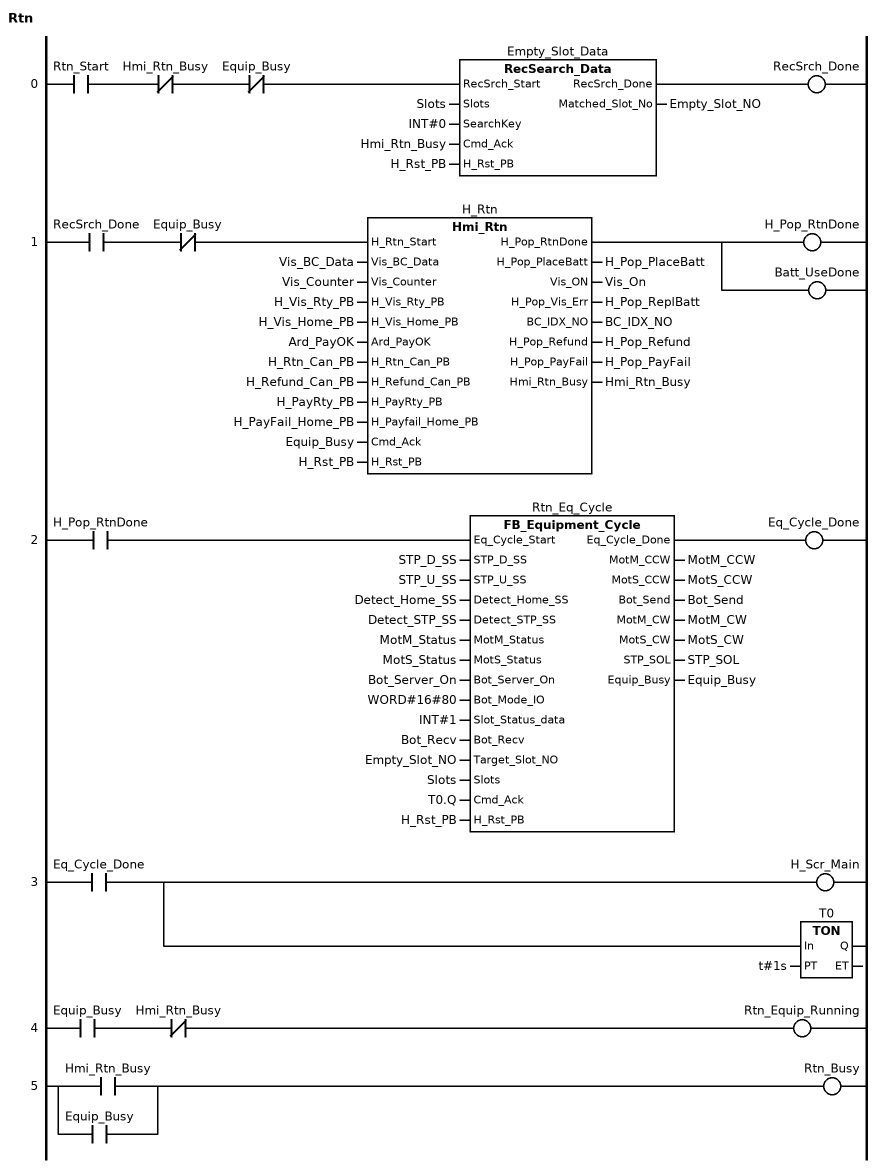
(* Rung 0 *)
Empty_Slot_Data(RecSrch_Start := Rtn_Start AND NOT Hmi_Rtn_Busy AND NOT Equip_Busy, Slots := Slots, SearchKey := INT#0, Cmd_Ack := Hmi_Rtn_Busy, H_Rst_PB := H_Rst_PB, Matched_Slot_No => Empty_Slot_NO);
RecSrch_Done := Empty_Slot_Data.RecSrch_Done;
(* Rung 1 *)
H_Rtn(H_Rtn_Start := RecSrch_Done AND NOT Equip_Busy, Vis_BC_Data := Vis_BC_Data, Vis_Counter := Vis_Counter, H_Vis_Rty_PB := H_Vis_Rty_PB, H_Vis_Home_PB := H_Vis_Home_PB, Ard_PayOK := Ard_PayOK, H_Rtn_Can_PB := H_Rtn_Can_PB, H_Refund_Can_PB := H_Refund_Can_PB, H_PayRty_PB := H_PayRty_PB, H_Payfail_Home_PB := H_PayFail_Home_PB, Cmd_Ack := Equip_Busy, H_Rst_PB := H_Rst_PB, H_Pop_PlaceBatt => H_Pop_PlaceBatt, Vis_ON => Vis_On, H_Pop_Vis_Err => H_Pop_ReplBatt, BC_IDX_NO => BC_IDX_NO, H_Pop_Refund => H_Pop_Refund, H_Pop_PayFail => H_Pop_PayFail, Hmi_Rtn_Busy => Hmi_Rtn_Busy);
_p1 := H_Rtn.H_Pop_RtnDone;
H_Pop_RtnDone := _p1;
Batt_UseDone := _p1;
(* Rung 2 *)
Rtn_Eq_Cycle(Eq_Cycle_Start := H_Pop_RtnDone, STP_D_SS := STP_D_SS, STP_U_SS := STP_U_SS, Detect_Home_SS := Detect_Home_SS, Detect_STP_SS := Detect_STP_SS, MotM_Status := MotM_Status, MotS_Status := MotS_Status, Bot_Server_On := Bot_Server_On, Bot_Mode_IO := WORD#16#80, Slot_Status_data := INT#1, Bot_Recv := Bot_Recv, Target_Slot_NO := Empty_Slot_NO, Slots := Slots, Cmd_Ack := T0.Q, H_Rst_PB := H_Rst_PB, MotM_CCW => MotM_CCW, MotS_CCW => MotS_CCW, Bot_Send => Bot_Send, MotM_CW => MotM_CW, MotS_CW => MotS_CW, STP_SOL => STP_SOL, Equip_Busy => Equip_Busy);
Eq_Cycle_Done := Rtn_Eq_Cycle.Eq_Cycle_Done;
(* Rung 3 *)
H_Scr_Main := Eq_Cycle_Done;
T0(In := Eq_Cycle_Done, PT := t#1s);
(* Rung 4 *)
Rtn_Equip_Running := Equip_Busy AND NOT Hmi_Rtn_Busy;
(* Rung 5 *)
Rtn_Busy := Hmi_Rtn_Busy OR Equip_Busy;
END_FUNCTION_BLOCK

FUNCTION_BLOCK RecMax_Data
VAR
    RecMax_SOC : UINT;
    RecMax_Slot_No : ARRAY[1..6] OF UINT;
    data : INT;
    W_RecMax_Pos : UINT;
    Status_Data : ARRAY[0..5] OF UINT;
    Match_Found : BOOL;
END_VAR
VAR_INPUT
    RecMax_Start : BOOL;
END_VAR
VAR_OUTPUT
    RecMax_Done : BOOL;
END_VAR
VAR_INPUT
    Slots : ARRAY[1..6] OF Slot_info;
END_VAR
VAR_OUTPUT
    Max_SOC : UINT;
    Max_Slot_NO : UINT;
END_VAR
VAR_INPUT
    Cmd_Ack : BOOL;
    H_Rst_PB : BOOL;
END_VAR
VAR
    _e1 : R_TRIG;
    _p2 : BOOL;
END_VAR
(* ladder, written here as Structured Text *)

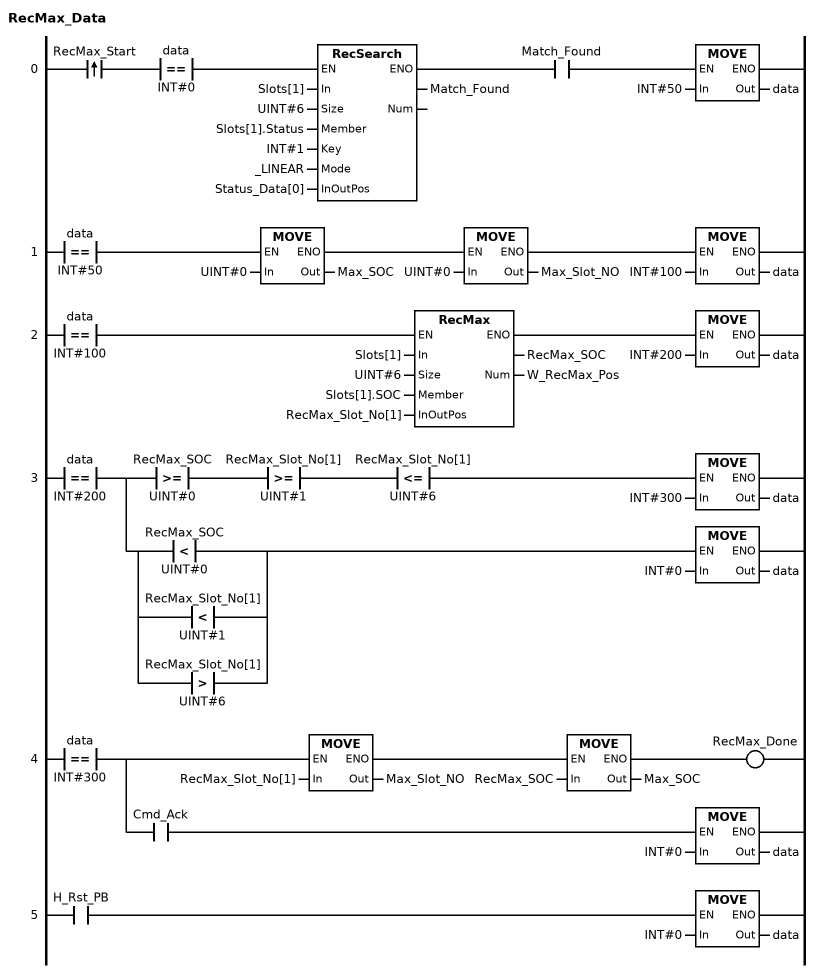
(* Rung 0 *)
_e1(CLK := RecMax_Start);
IF _e1.Q AND (data = INT#0) THEN
    Match_Found := RecSearch(In := Slots[1], Size := UINT#6, Member := Slots[1].Status, Key := INT#1, Mode := _LINEAR, InOutPos := Status_Data[0]);
END_IF;
IF _e1.Q AND (data = INT#0) AND Match_Found THEN data := INT#50; END_IF;
(* Rung 1 *)
IF data = INT#50 THEN
    Max_SOC := UINT#0;
    Max_Slot_NO := UINT#0;
    data := INT#100;
END_IF;
(* Rung 2 *)
IF data = INT#100 THEN
    RecMax_SOC := RecMax(In := Slots[1], Size := UINT#6, Member := Slots[1].SOC, InOutPos := RecMax_Slot_No[1], Num => W_RecMax_Pos);
    data := INT#200;
END_IF;
(* Rung 3 *)
_p2 := data = INT#200;
IF (data = INT#200) AND (RecMax_SOC >= UINT#0) AND (RecMax_Slot_No[1] >= UINT#1) AND (RecMax_Slot_No[1] <= UINT#6) THEN
    data := INT#300;
END_IF;
IF _p2 AND ((RecMax_SOC < UINT#0) OR (RecMax_Slot_No[1] < UINT#1) OR (RecMax_Slot_No[1] > UINT#6)) THEN
    data := INT#0;
END_IF;
(* Rung 4 *)
IF data = INT#300 THEN
    Max_Slot_NO := RecMax_Slot_No[1];
    Max_SOC := RecMax_SOC;
END_IF;
RecMax_Done := data = INT#300;
IF (data = INT#300) AND Cmd_Ack THEN data := INT#0; END_IF;
(* Rung 5 *)
IF H_Rst_PB THEN data := INT#0; END_IF;
END_FUNCTION_BLOCK

FUNCTION_BLOCK Hmi_Rtn
VAR
    data : INT;
    T0 : TON;
    Vis_Rtn : Vision;
    Vis_Busy : BOOL;
    T1 : TON;
    T2 : TON;
END_VAR
VAR_INPUT
    H_Rtn_Start : BOOL;
END_VAR
VAR_OUTPUT
    H_Pop_RtnDone : BOOL;
    H_Pop_PlaceBatt : BOOL;
    Vis_ON : BOOL;
END_VAR
VAR_INPUT
    Vis_BC_Data : DINT;
    Vis_Counter : DINT;
    H_Vis_Rty_PB : BOOL;
    H_Vis_Home_PB : BOOL;
END_VAR
VAR_OUTPUT
    H_Pop_Vis_Err : BOOL;
    BC_IDX_NO : DINT;
END_VAR
VAR_INPUT
    Ard_PayOK : BOOL;
END_VAR
VAR_OUTPUT
    H_Pop_Refund : BOOL;
END_VAR
VAR_INPUT
    H_Rtn_Can_PB : BOOL;
    H_Refund_Can_PB : BOOL;
    H_PayRty_PB : BOOL;
    H_Payfail_Home_PB : BOOL;
    Cmd_Ack : BOOL;
END_VAR
VAR_OUTPUT
    H_Pop_PayFail : BOOL;
    Hmi_Rtn_Busy : BOOL;
END_VAR
VAR_INPUT
    H_Rst_PB : BOOL;
END_VAR
VAR
    _e1 : R_TRIG;
    _p2 : BOOL;
    _p3 : BOOL;
    _p4 : BOOL;
    _p5 : BOOL;
END_VAR
(* ladder, written here as Structured Text *)

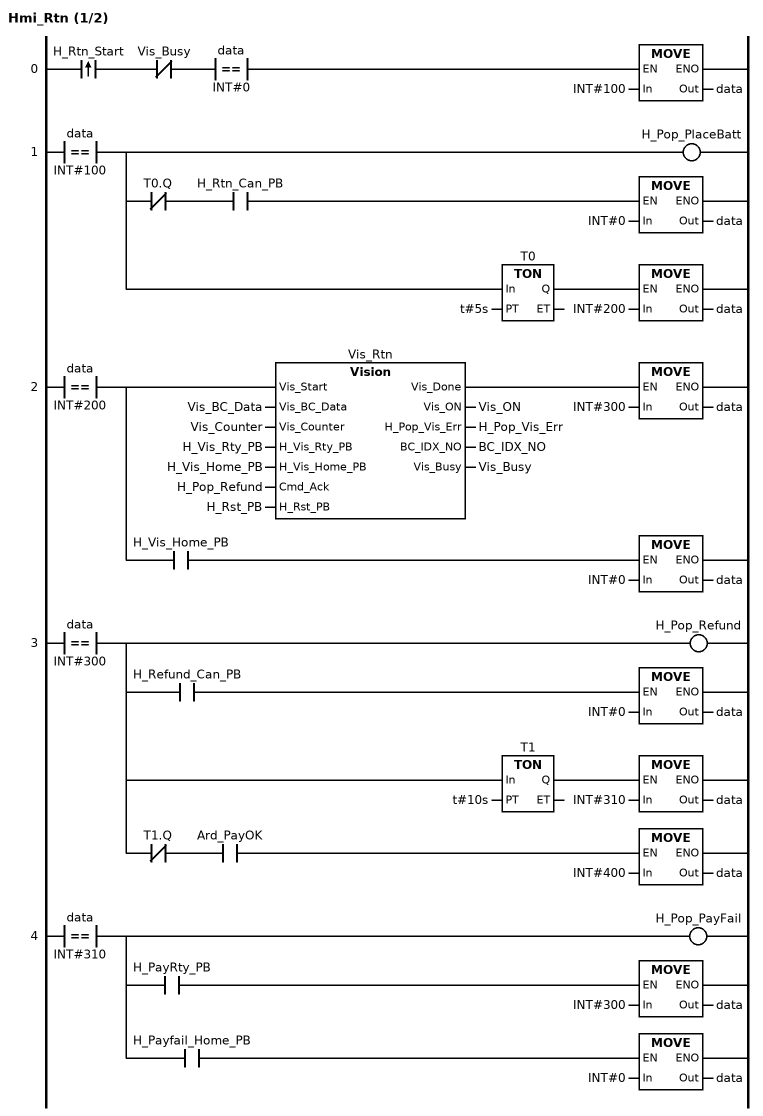
(* Rung 0 *)
_e1(CLK := H_Rtn_Start);
IF _e1.Q AND NOT Vis_Busy AND (data = INT#0) THEN data := INT#100; END_IF;
(* Rung 1 *)
H_Pop_PlaceBatt := data = INT#100;
_p2 := data = INT#100;
IF (data = INT#100) AND NOT T0.Q AND H_Rtn_Can_PB THEN data := INT#0; END_IF;
T0(In := _p2, PT := t#5s);
IF T0.Q THEN data := INT#200; END_IF;
(* Rung 2 *)
Vis_Rtn(Vis_Start := data = INT#200, Vis_BC_Data := Vis_BC_Data, Vis_Counter := Vis_Counter, H_Vis_Rty_PB := H_Vis_Rty_PB, H_Vis_Home_PB := H_Vis_Home_PB, Cmd_Ack := H_Pop_Refund, H_Rst_PB := H_Rst_PB, Vis_ON => Vis_ON, H_Pop_Vis_Err => H_Pop_Vis_Err, BC_IDX_NO => BC_IDX_NO, Vis_Busy => Vis_Busy);
_p3 := data = INT#200;
IF Vis_Rtn.Vis_Done THEN data := INT#300; END_IF;
IF _p3 AND H_Vis_Home_PB THEN data := INT#0; END_IF;
(* Rung 3 *)
H_Pop_Refund := data = INT#300;
_p4 := data = INT#300;
IF (data = INT#300) AND H_Refund_Can_PB THEN data := INT#0; END_IF;
T1(In := _p4, PT := t#10s);
IF T1.Q THEN data := INT#310; END_IF;
IF _p4 AND NOT T1.Q AND Ard_PayOK THEN data := INT#400; END_IF;
(* Rung 4 *)
H_Pop_PayFail := data = INT#310;
_p5 := data = INT#310;
IF (data = INT#310) AND H_PayRty_PB THEN data := INT#300; END_IF;
IF _p5 AND H_Payfail_Home_PB THEN data := INT#0; END_IF;

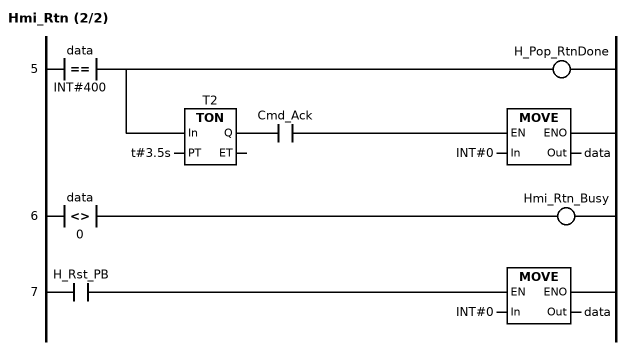
(* Rung 5 *)
H_Pop_RtnDone := data = INT#400;
T2(In := data = INT#400, PT := t#3.5s);
IF T2.Q AND Cmd_Ack THEN data := INT#0; END_IF;
(* Rung 6 *)
Hmi_Rtn_Busy := data <> 0;
(* Rung 7 *)
IF H_Rst_PB THEN data := INT#0; END_IF;
END_FUNCTION_BLOCK

FUNCTION_BLOCK RecSearch_Data
VAR
    MatchFound : BOOL;
    data : INT;
    RecSrch_data : ARRAY[1..6] OF UINT;
    W_RecSrch_Pos : UINT;
END_VAR
VAR_INPUT
    RecSrch_Start : BOOL;
END_VAR
VAR_OUTPUT
    RecSrch_Done : BOOL;
END_VAR
VAR_INPUT
    Slots : ARRAY[1..6] OF Slot_info;
    SearchKey : INT;
END_VAR
VAR_OUTPUT
    Matched_Slot_No : UINT;
END_VAR
VAR_INPUT
    Cmd_Ack : BOOL;
    H_Rst_PB : BOOL;
END_VAR
VAR
    _p1 : BOOL;
END_VAR
(* ladder, written here as Structured Text *)

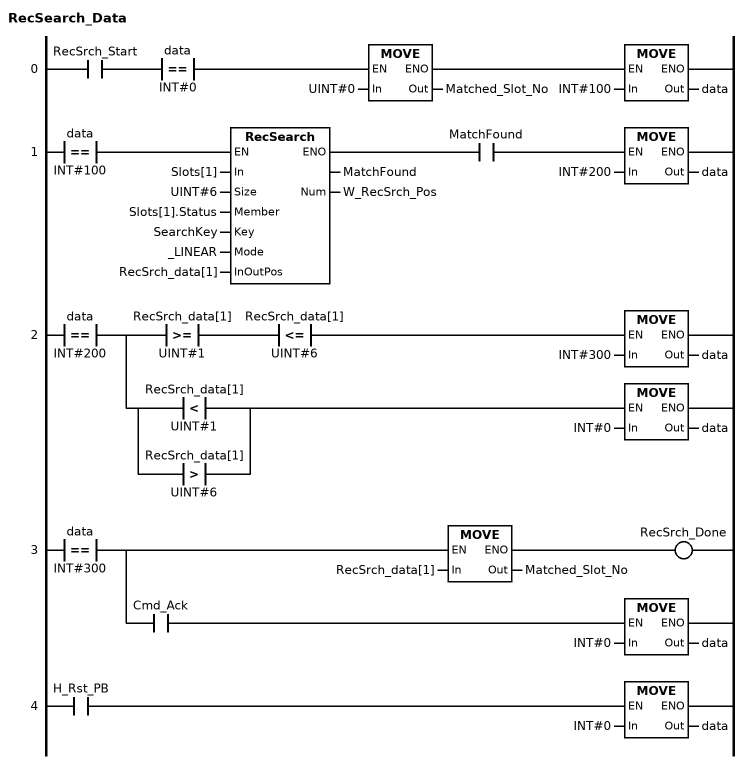
(* Rung 0 *)
IF RecSrch_Start AND (data = INT#0) THEN
    Matched_Slot_No := UINT#0;
    data := INT#100;
END_IF;
(* Rung 1 *)
IF data = INT#100 THEN
    MatchFound := RecSearch(In := Slots[1], Size := UINT#6, Member := Slots[1].Status, Key := SearchKey, Mode := _LINEAR, InOutPos := RecSrch_data[1], Num => W_RecSrch_Pos);
END_IF;
IF (data = INT#100) AND MatchFound THEN data := INT#200; END_IF;
(* Rung 2 *)
_p1 := data = INT#200;
IF (data = INT#200) AND (RecSrch_data[1] >= UINT#1) AND (RecSrch_data[1] <= UINT#6) THEN
    data := INT#300;
END_IF;
IF _p1 AND ((RecSrch_data[1] < UINT#1) OR (RecSrch_data[1] > UINT#6)) THEN data := INT#0; END_IF;
(* Rung 3 *)
IF data = INT#300 THEN Matched_Slot_No := RecSrch_data[1]; END_IF;
RecSrch_Done := data = INT#300;
IF (data = INT#300) AND Cmd_Ack THEN data := INT#0; END_IF;
(* Rung 4 *)
IF H_Rst_PB THEN data := INT#0; END_IF;
END_FUNCTION_BLOCK

FUNCTION_BLOCK FB_Equipment_Cycle
VAR
    MPS_Home_To_Bot : MPS;
    Bot_Done : BOOL;
    MPS_Done : BOOL;
    Rent_Robot : Robot_Move;
    MPS_Bot_To_Home : MPS;
    STP_D_SOL : BOOL;
    STP_U_SOL : BOOL;
    Robot_Busy : BOOL;
    Mps_Busy : ARRAY[0..1] OF BOOL;
    Bot_Clear : BOOL;
    Mps_Home_Done : BOOL;
END_VAR
VAR_INPUT
    Eq_Cycle_Start : BOOL;
END_VAR
VAR_OUTPUT
    Eq_Cycle_Done : BOOL;
END_VAR
VAR_INPUT
    STP_D_SS : BOOL;
    STP_U_SS : BOOL;
    Detect_Home_SS : BOOL;
    Detect_STP_SS : BOOL;
END_VAR
VAR_OUTPUT
    MotM_CCW : BOOL;
    MotS_CCW : BOOL;
END_VAR
VAR_INPUT
    MotM_Status : WORD;
    MotS_Status : WORD;
    Bot_Server_On : BOOL;
    Bot_Mode_IO : WORD;
    Slot_Status_data : INT;
END_VAR
VAR_OUTPUT
    Bot_Send : S_RobotIO;
END_VAR
VAR_INPUT
    Bot_Recv : S_RobotIO;
    Target_Slot_NO : UINT;
END_VAR
VAR_OUTPUT
    MotM_CW : BOOL;
END_VAR
VAR_IN_OUT
    Slots : ARRAY[1..6] OF Slot_info;
END_VAR
VAR_INPUT
    Cmd_Ack : BOOL;
END_VAR
VAR_OUTPUT
    MotS_CW : BOOL;
    STP_SOL : BOOL;
    Equip_Busy : BOOL;
END_VAR
VAR_INPUT
    H_Rst_PB : BOOL;
END_VAR
VAR
    _p1 : BOOL;
    _p2 : BOOL;
END_VAR
(* ladder, written here as Structured Text *)

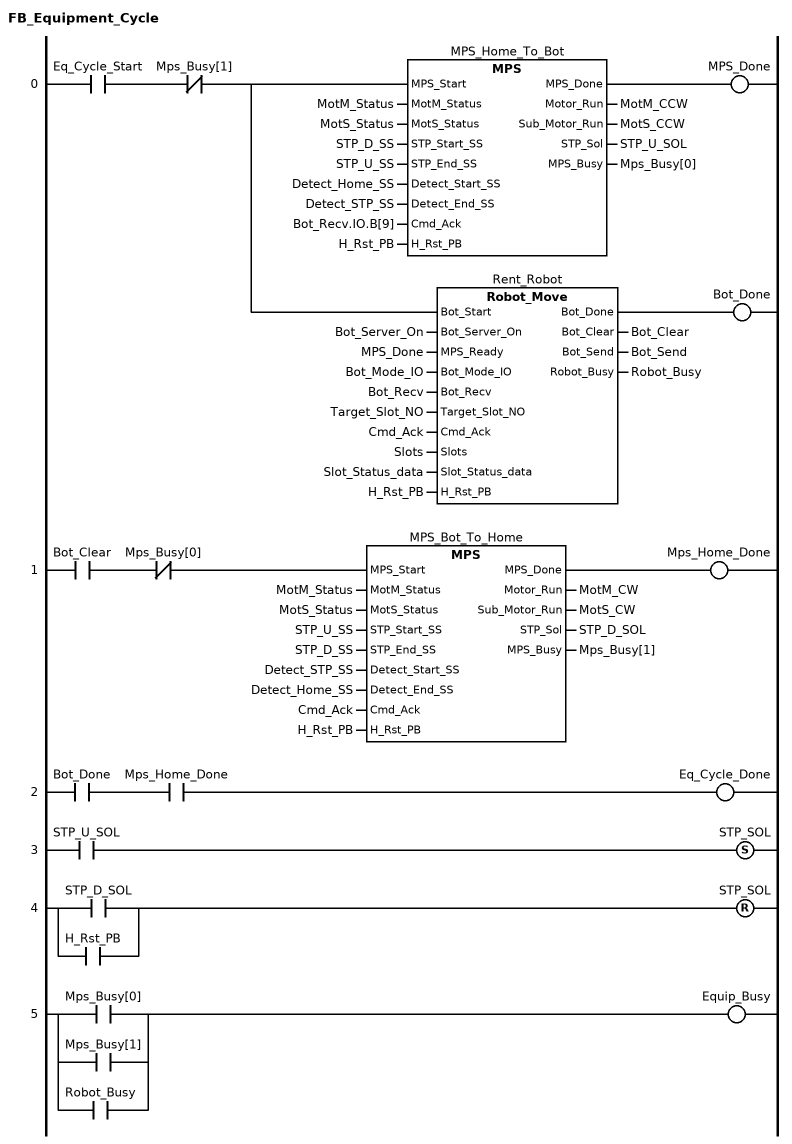
(* Rung 0 *)
_p1 := Eq_Cycle_Start AND NOT Mps_Busy[1];
MPS_Home_To_Bot(MPS_Start := _p1, MotM_Status := MotM_Status, MotS_Status := MotS_Status, STP_Start_SS := STP_D_SS, STP_End_SS := STP_U_SS, Detect_Start_SS := Detect_Home_SS, Detect_End_SS := Detect_STP_SS, Cmd_Ack := Bot_Recv.IO.B[9], H_Rst_PB := H_Rst_PB, Motor_Run => MotM_CCW, Sub_Motor_Run => MotS_CCW, STP_Sol => STP_U_SOL, MPS_Busy => Mps_Busy[0]);
MPS_Done := MPS_Home_To_Bot.MPS_Done;
Rent_Robot(Bot_Start := _p1, Bot_Server_On := Bot_Server_On, MPS_Ready := MPS_Done, Bot_Mode_IO := Bot_Mode_IO, Bot_Recv := Bot_Recv, Target_Slot_NO := Target_Slot_NO, Cmd_Ack := Cmd_Ack, Slots := Slots, Slot_Status_data := Slot_Status_data, H_Rst_PB := H_Rst_PB, Bot_Clear => Bot_Clear, Bot_Send => Bot_Send, Robot_Busy => Robot_Busy);
Bot_Done := Rent_Robot.Bot_Done;
(* Rung 1 *)
_p2 := Bot_Clear AND NOT Mps_Busy[0];
MPS_Bot_To_Home(MPS_Start := _p2, MotM_Status := MotM_Status, MotS_Status := MotS_Status, STP_Start_SS := STP_U_SS, STP_End_SS := STP_D_SS, Detect_Start_SS := Detect_STP_SS, Detect_End_SS := Detect_Home_SS, Cmd_Ack := Cmd_Ack, H_Rst_PB := H_Rst_PB, Motor_Run => MotM_CW, Sub_Motor_Run => MotS_CW, STP_Sol => STP_D_SOL, MPS_Busy => Mps_Busy[1]);
Mps_Home_Done := MPS_Bot_To_Home.MPS_Done;
(* Rung 2 *)
Eq_Cycle_Done := Bot_Done AND Mps_Home_Done;
(* Rung 3 *)
IF STP_U_SOL THEN STP_SOL := TRUE; END_IF;
(* Rung 4 *)
IF STP_D_SOL OR H_Rst_PB THEN STP_SOL := FALSE; END_IF;
(* Rung 5 *)
Equip_Busy := Mps_Busy[0] OR Mps_Busy[1] OR Robot_Busy;
END_FUNCTION_BLOCK

FUNCTION_BLOCK NG
VAR
    W_RecSrch_Pos : ARRAY[0..5] OF UINT;
    data : INT;
    NG_RecSrch : RecSearch_Data;
    NGBatt_Slot_No : UINT;
    Bot_Done : BOOL;
    T0 : TON;
    Bot_MV_BattNG : Bot_Move_NGBatt;
END_VAR
VAR_INPUT
    NG_Start : BOOL;
END_VAR
VAR_IN_OUT
    Slots : ARRAY[1..6] OF Slot_info;
END_VAR
VAR_INPUT
    Bot_Server_On : BOOL;
END_VAR
VAR_OUTPUT
    H_Pop_BattNG_Running : BOOL;
    H_Scr_Main : BOOL;
END_VAR
VAR_INPUT
    Bot_Recv : S_RobotIO;
END_VAR
VAR_OUTPUT
    Bot_Send : S_RobotIO;
    RecSrch_Done : BOOL;
    NG_Busy : BOOL;
END_VAR
VAR_INPUT
    H_Rst_PB : BOOL;
END_VAR
(* ladder, written here as Structured Text *)

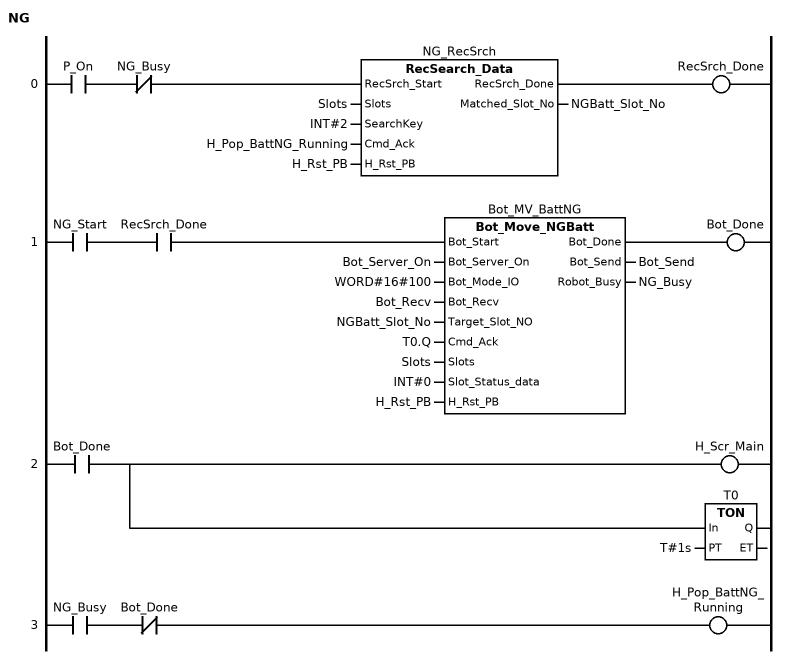
(* Rung 0 *)
NG_RecSrch(RecSrch_Start := P_On AND NOT NG_Busy, Slots := Slots, SearchKey := INT#2, Cmd_Ack := H_Pop_BattNG_Running, H_Rst_PB := H_Rst_PB, Matched_Slot_No => NGBatt_Slot_No);
RecSrch_Done := NG_RecSrch.RecSrch_Done;
(* Rung 1 *)
Bot_MV_BattNG(Bot_Start := NG_Start AND RecSrch_Done, Bot_Server_On := Bot_Server_On, Bot_Mode_IO := WORD#16#100, Bot_Recv := Bot_Recv, Target_Slot_NO := NGBatt_Slot_No, Cmd_Ack := T0.Q, Slots := Slots, Slot_Status_data := INT#0, H_Rst_PB := H_Rst_PB, Bot_Send => Bot_Send, Robot_Busy => NG_Busy);
Bot_Done := Bot_MV_BattNG.Bot_Done;
(* Rung 2 *)
H_Scr_Main := Bot_Done;
T0(In := Bot_Done, PT := T#1s);
(* Rung 3 *)
H_Pop_BattNG_Running := NG_Busy AND NOT Bot_Done;
END_FUNCTION_BLOCK

FUNCTION_BLOCK Bot_Move_NGBatt
VAR
    Cmd_Base : WORD;
    data : INT;
END_VAR
VAR_INPUT
    Bot_Start : BOOL;
END_VAR
VAR_OUTPUT
    Bot_Done : BOOL;
END_VAR
VAR_INPUT
    Bot_Server_On : BOOL;
    Bot_Mode_IO : WORD;
    Bot_Recv : S_RobotIO;
    Target_Slot_NO : UINT;
END_VAR
VAR_OUTPUT
    Bot_Send : S_RobotIO;
END_VAR
VAR_INPUT
    Cmd_Ack : BOOL;
END_VAR
VAR_IN_OUT
    Slots : ARRAY[1..6] OF Slot_info;
END_VAR
VAR_INPUT
    Slot_Status_data : INT;
END_VAR
VAR_OUTPUT
    Robot_Busy : BOOL;
END_VAR
VAR_INPUT
    H_Rst_PB : BOOL;
END_VAR
VAR
    _p1 : BOOL;
END_VAR
(* ladder, written here as Structured Text *)

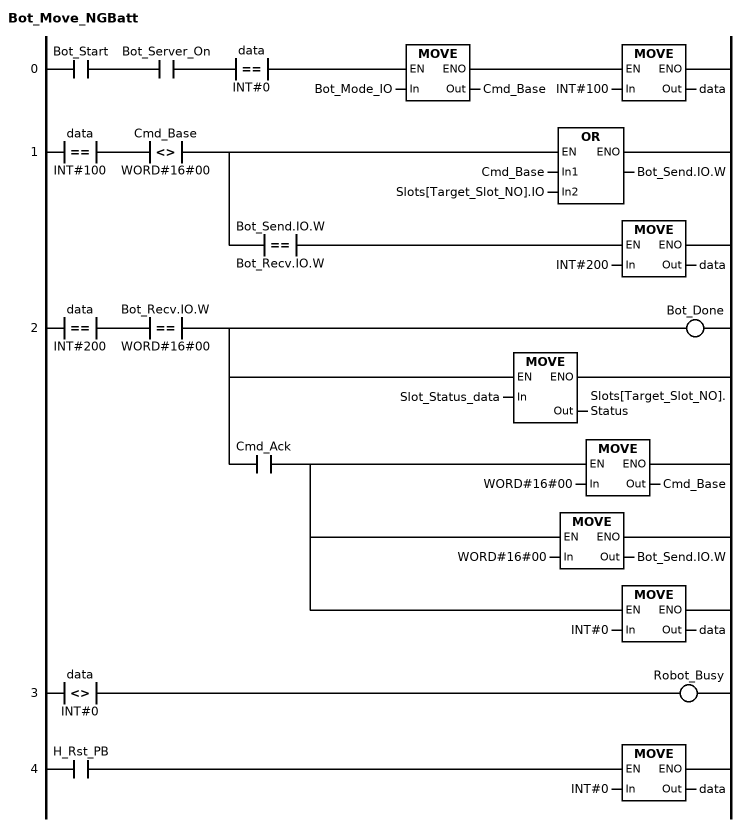
(* Rung 0 *)
IF Bot_Start AND Bot_Server_On AND (data = INT#0) THEN
    Cmd_Base := Bot_Mode_IO;
    data := INT#100;
END_IF;
(* Rung 1 *)
IF (data = INT#100) AND (Cmd_Base <> WORD#16#00) THEN
    Bot_Send.IO.W := Cmd_Base OR Slots[Target_Slot_NO].IO;
END_IF;
IF (data = INT#100) AND (Cmd_Base <> WORD#16#00) AND (Bot_Send.IO.W = Bot_Recv.IO.W) THEN
    data := INT#200;
END_IF;
(* Rung 2 *)
_p1 := (data = INT#200) AND (Bot_Recv.IO.W = WORD#16#00);
Bot_Done := _p1;
IF _p1 THEN Slots[Target_Slot_NO].Status := Slot_Status_data; END_IF;
IF _p1 AND Cmd_Ack THEN
    Cmd_Base := WORD#16#00;
    Bot_Send.IO.W := WORD#16#00;
    data := INT#0;
END_IF;
(* Rung 3 *)
Robot_Busy := data <> INT#0;
(* Rung 4 *)
IF H_Rst_PB THEN data := INT#0; END_IF;
END_FUNCTION_BLOCK

FUNCTION_BLOCK FB_Batt_Process
VAR
    Batt_Rtn : Rtn;
    Batt_Rent : Rent;
    Batt_NG : NG;
    Mot1_CCW : ARRAY[0..1] OF BOOL;
    Mot1_CW : ARRAY[0..1] OF BOOL;
    Mot2_CCW : ARRAY[0..1] OF BOOL;
    Mot2_CW : ARRAY[0..1] OF BOOL;
    Bot_Send_Data : ARRAY[0..2] OF S_RobotIO;
    Stopper_SOL : ARRAY[0..1] OF BOOL;
    Vision_On : ARRAY[0..1] OF BOOL;
    Rent_BC_IDX : DINT;
    H_Main_Screen : ARRAY[0..2] OF BOOL;
    Rent_Busy : BOOL;
    Rtn_Busy : BOOL;
    NG_Busy : BOOL;
    Batt_UseStart : BOOL;
    Batt_UseDone : BOOL;
END_VAR
VAR RETAIN
    Batt_IsUse : ARRAY[1..6] OF BOOL;
END_VAR
VAR
    Bot_Recv_Data : S_RobotIO;
    Batt_NG_Running : BOOL;
    MotM_CW : BOOL;
    MotM_CCW : BOOL;
    MotS_CW : BOOL;
    MotS_CCW : BOOL;
    BC_NO_MFC : WORD;
    Hmi_Pop_PayFail : ARRAY[0..1] OF BOOL;
    Rtn_Equip_Running : BOOL;
END_VAR
VAR RETAIN
    Batt_RentTime : ARRAY[1..6] OF DATE_AND_TIME;
END_VAR
VAR
    NG_Ready : BOOL;
    UseSec : DINT;
    i : INT;
END_VAR
VAR_INPUT
    H_Rent_PB : BOOL;
    Ard_PayOK : BOOL;
    H_Card_Can_PB : BOOL;
    H_LowBatt_OK_PB : BOOL;
    H_LowBatt_Can_PB : BOOL;
    MotM_Status : WORD;
    MotS_Status : WORD;
END_VAR
VAR_IN_OUT
    Slots : ARRAY[1..6] OF Slot_info;
END_VAR
VAR_INPUT
    STP_D_SS : BOOL;
    STP_U_SS : BOOL;
    Detect_Home_SS : BOOL;
    Detect_STP_SS : BOOL;
    Bot_Server_ON : BOOL;
    Bot_Recv : S_RobotIO;
    H_Rtn_PB : BOOL;
    H_Vis_Rty_PB : BOOL;
    H_Vis_Home_PB : BOOL;
    Vis_BC_Data : DINT;
    Vis_Counter_Data : DINT;
    H_Rtn_Can_PB : BOOL;
    H_Refund_Can_PB : BOOL;
    H_PayRty_PB : BOOL;
    H_PayFail_Home_PB : BOOL;
END_VAR
VAR_OUTPUT
    H_Pop_Card : BOOL;
    H_Pop_Wait_Rent : BOOL;
    H_Pop_LowBatt : BOOL;
    MotM_MV : WORD;
    MotS_MV : WORD;
    H_Pop_ContAdmin : BOOL;
    H_Pop_PayFail : BOOL;
    H_Pop_Rent_Done : BOOL;
    H_Pop_Place_Batt : BOOL;
    H_Pop_ReplBatt : BOOL;
    H_Pop_Refund : BOOL;
    H_Pop_RtnDone : BOOL;
    H_Pop_BattNG_Running : BOOL;
    Bot_Send : S_RobotIO;
    STP_SOL : BOOL;
    Vision_Trigger_On : BOOL;
    H_Scr_Main : BOOL;
    Rtn_BC_IDX : DINT;
    Batt_UseTime : ARRAY[1..6] OF TIME;
    Batt_UseDisp : ARRAY[1..6] OF DINT;
    Max_SOC : UINT;
    Batt_Refund : LINT;
    Batt_UseFee : LINT;
END_VAR
VAR_INPUT
    H_Rst_PB : BOOL;
END_VAR
VAR_EXTERNAL
    MFC_HR : ARRAY[0..99] OF WORD;
END_VAR
VAR_EXTERNAL CONSTANT
    _CurrentTime : DATE_AND_TIME;
END_VAR
VAR
    _e1 : R_TRIG;
    _e2 : R_TRIG;
    _e3 : R_TRIG;
END_VAR
(* ladder, written here as Structured Text *)

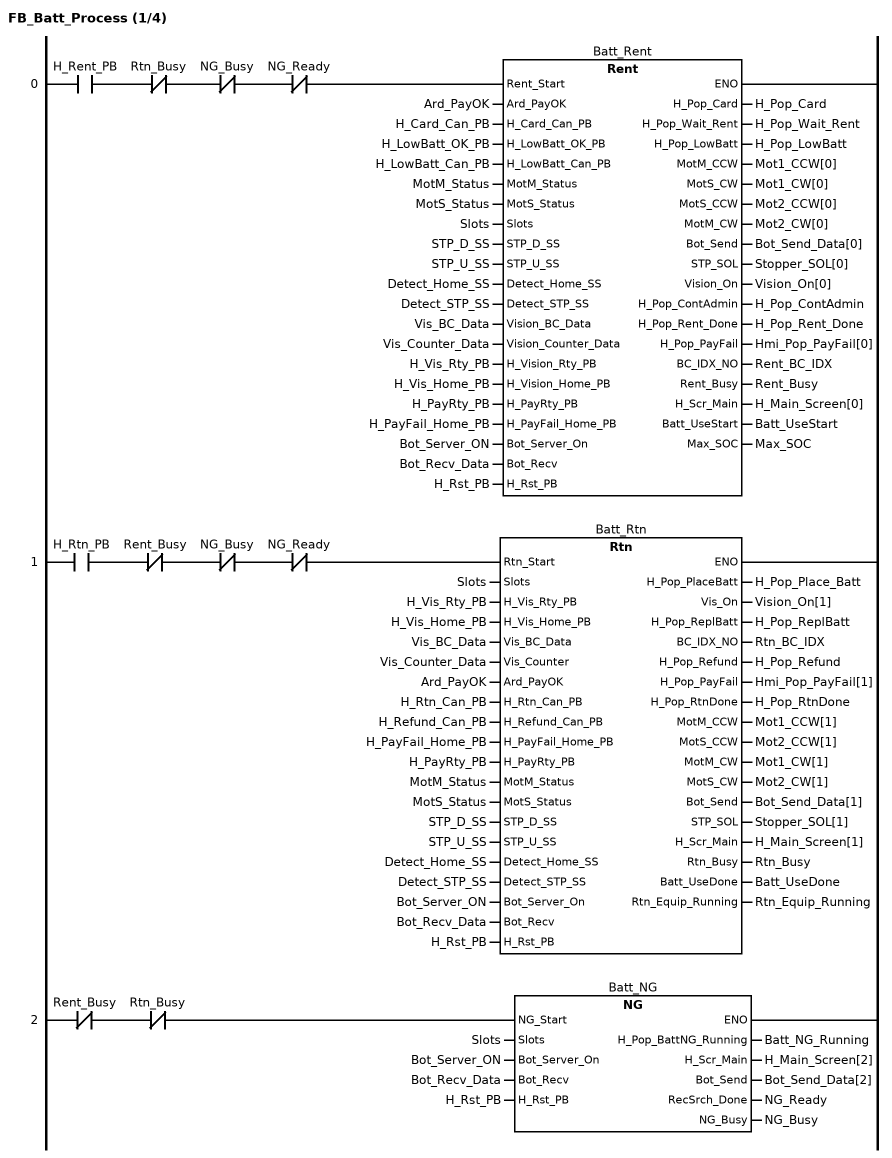
(* Rung 0 *)
Batt_Rent(Rent_Start := H_Rent_PB AND NOT Rtn_Busy AND NOT NG_Busy AND NOT NG_Ready, Ard_PayOK := Ard_PayOK, H_Card_Can_PB := H_Card_Can_PB, H_LowBatt_OK_PB := H_LowBatt_OK_PB, H_LowBatt_Can_PB := H_LowBatt_Can_PB, MotM_Status := MotM_Status, MotS_Status := MotS_Status, Slots := Slots, STP_D_SS := STP_D_SS, STP_U_SS := STP_U_SS, Detect_Home_SS := Detect_Home_SS, Detect_STP_SS := Detect_STP_SS, Vision_BC_Data := Vis_BC_Data, Vision_Counter_Data := Vis_Counter_Data, H_Vision_Rty_PB := H_Vis_Rty_PB, H_Vision_Home_PB := H_Vis_Home_PB, H_PayRty_PB := H_PayRty_PB, H_PayFail_Home_PB := H_PayFail_Home_PB, Bot_Server_On := Bot_Server_ON, Bot_Recv := Bot_Recv_Data, H_Rst_PB := H_Rst_PB, H_Pop_Card => H_Pop_Card, H_Pop_Wait_Rent => H_Pop_Wait_Rent, H_Pop_LowBatt => H_Pop_LowBatt, MotM_CCW => Mot1_CCW[0], MotS_CW => Mot1_CW[0], MotS_CCW => Mot2_CCW[0], MotM_CW => Mot2_CW[0], Bot_Send => Bot_Send_Data[0], STP_SOL => Stopper_SOL[0], Vision_On => Vision_On[0], H_Pop_ContAdmin => H_Pop_ContAdmin, H_Pop_Rent_Done => H_Pop_Rent_Done, H_Pop_PayFail => Hmi_Pop_PayFail[0], BC_IDX_NO => Rent_BC_IDX, Rent_Busy => Rent_Busy, H_Scr_Main => H_Main_Screen[0], Batt_UseStart => Batt_UseStart, Max_SOC => Max_SOC);
(* Rung 1 *)
Batt_Rtn(Rtn_Start := H_Rtn_PB AND NOT Rent_Busy AND NOT NG_Busy AND NOT NG_Ready, Slots := Slots, H_Vis_Rty_PB := H_Vis_Rty_PB, H_Vis_Home_PB := H_Vis_Home_PB, Vis_BC_Data := Vis_BC_Data, Vis_Counter := Vis_Counter_Data, Ard_PayOK := Ard_PayOK, H_Rtn_Can_PB := H_Rtn_Can_PB, H_Refund_Can_PB := H_Refund_Can_PB, H_PayFail_Home_PB := H_PayFail_Home_PB, H_PayRty_PB := H_PayRty_PB, MotM_Status := MotM_Status, MotS_Status := MotS_Status, STP_D_SS := STP_D_SS, STP_U_SS := STP_U_SS, Detect_Home_SS := Detect_Home_SS, Detect_STP_SS := Detect_STP_SS, Bot_Server_On := Bot_Server_ON, Bot_Recv := Bot_Recv_Data, H_Rst_PB := H_Rst_PB, H_Pop_PlaceBatt => H_Pop_Place_Batt, Vis_On => Vision_On[1], H_Pop_ReplBatt => H_Pop_ReplBatt, BC_IDX_NO => Rtn_BC_IDX, H_Pop_Refund => H_Pop_Refund, H_Pop_PayFail => Hmi_Pop_PayFail[1], H_Pop_RtnDone => H_Pop_RtnDone, MotM_CCW => Mot1_CCW[1], MotS_CCW => Mot2_CCW[1], MotM_CW => Mot1_CW[1], MotS_CW => Mot2_CW[1], Bot_Send => Bot_Send_Data[1], STP_SOL => Stopper_SOL[1], H_Scr_Main => H_Main_Screen[1], Rtn_Busy => Rtn_Busy, Batt_UseDone => Batt_UseDone, Rtn_Equip_Running => Rtn_Equip_Running);
(* Rung 2 *)
Batt_NG(NG_Start := NOT Rent_Busy AND NOT Rtn_Busy, Slots := Slots, Bot_Server_On := Bot_Server_ON, Bot_Recv := Bot_Recv_Data, H_Rst_PB := H_Rst_PB, H_Pop_BattNG_Running => Batt_NG_Running, H_Scr_Main => H_Main_Screen[2], Bot_Send => Bot_Send_Data[2], RecSrch_Done => NG_Ready, NG_Busy => NG_Busy);

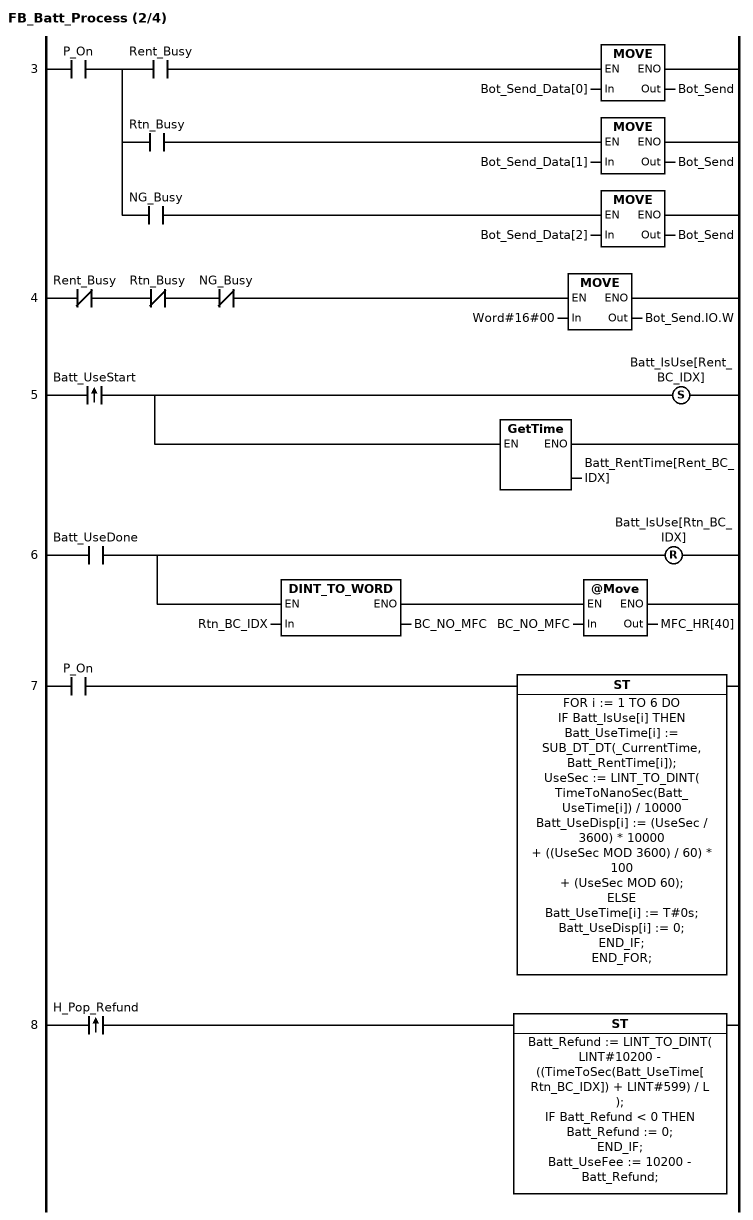
(* Rung 3 *)
IF P_On AND Rent_Busy THEN Bot_Send := Bot_Send_Data[0]; END_IF;
IF P_On AND Rtn_Busy THEN Bot_Send := Bot_Send_Data[1]; END_IF;
IF P_On AND NG_Busy THEN Bot_Send := Bot_Send_Data[2]; END_IF;
(* Rung 4 *)
IF NOT Rent_Busy AND NOT Rtn_Busy AND NOT NG_Busy THEN Bot_Send.IO.W := Word#16#00; END_IF;
(* Rung 5 *)
_e1(CLK := Batt_UseStart);
IF _e1.Q THEN
    Batt_IsUse[Rent_BC_IDX] := TRUE;
    Batt_RentTime[Rent_BC_IDX] := GetTime();
END_IF;
(* Rung 6 *)
IF Batt_UseDone THEN
    Batt_IsUse[Rtn_BC_IDX] := FALSE;
    BC_NO_MFC := DINT_TO_WORD(In := Rtn_BC_IDX);
END_IF;
_e2(CLK := Batt_UseDone);
IF _e2.Q THEN MFC_HR[40] := BC_NO_MFC; END_IF;
(* Rung 7 *)
IF P_On THEN
    FOR i := 1 TO 6 DO
        IF Batt_IsUse[i] THEN
            Batt_UseTime[i] := SUB_DT_DT(_CurrentTime, Batt_RentTime[i]);
            UseSec := LINT_TO_DINT( TimeToNanoSec(Batt_UseTime[i]) / 1000000000 );
            Batt_UseDisp[i] := (UseSec / 3600) * 10000
                             + ((UseSec MOD 3600) / 60) * 100
                             + (UseSec MOD 60);
        ELSE
            Batt_UseTime[i] := T#0s;      
            Batt_UseDisp[i] := 0;
        END_IF;
    END_FOR;
END_IF;
(* Rung 8 *)
_e3(CLK := H_Pop_Refund);
IF _e3.Q THEN
    Batt_Refund := LINT_TO_DINT(
        LINT#10200 - ((TimeToSec(Batt_UseTime[Rtn_BC_IDX]) + LINT#599) / LINT#600) * LINT#200
    );
    
    IF Batt_Refund < 0 THEN
        Batt_Refund := 0;
    END_IF;
    
    Batt_UseFee := 10200 - Batt_Refund;
END_IF;

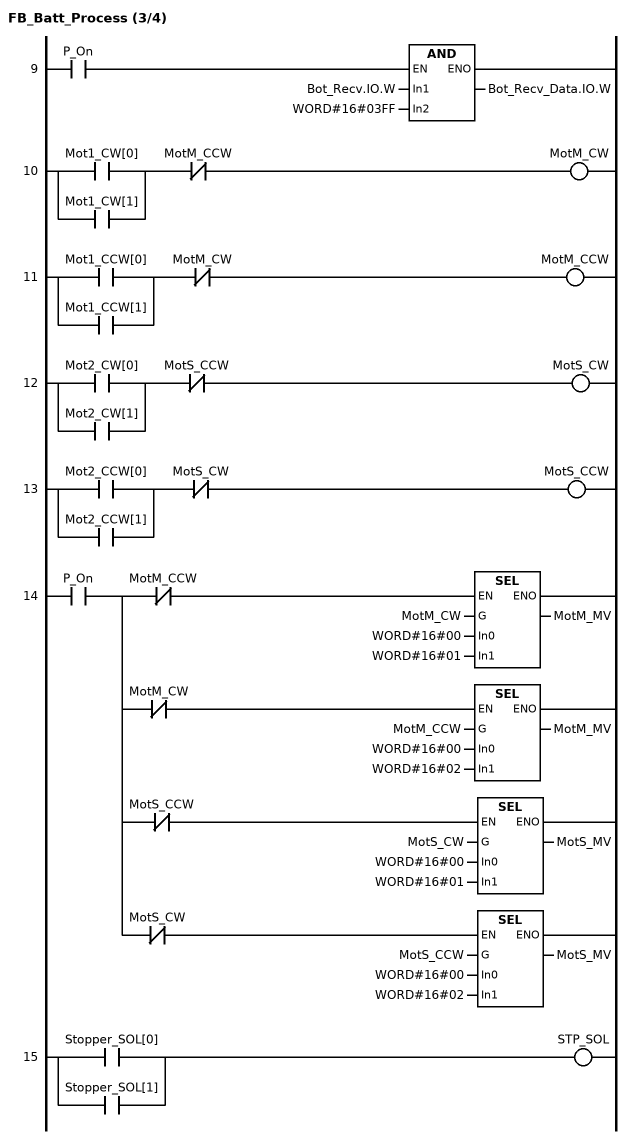
(* Rung 9 *)
IF P_On THEN Bot_Recv_Data.IO.W := Bot_Recv.IO.W AND WORD#16#03FF; END_IF;
(* Rung 10 *)
MotM_CW := (Mot1_CW[0] OR Mot1_CW[1]) AND NOT MotM_CCW;
(* Rung 11 *)
MotM_CCW := (Mot1_CCW[0] OR Mot1_CCW[1]) AND NOT MotM_CW;
(* Rung 12 *)
MotS_CW := (Mot2_CW[0] OR Mot2_CW[1]) AND NOT MotS_CCW;
(* Rung 13 *)
MotS_CCW := (Mot2_CCW[0] OR Mot2_CCW[1]) AND NOT MotS_CW;
(* Rung 14 *)
IF P_On AND NOT MotM_CCW THEN MotM_MV := SEL(G := MotM_CW, In0 := WORD#16#00, In1 := WORD#16#01); END_IF;
IF P_On AND NOT MotM_CW THEN MotM_MV := SEL(G := MotM_CCW, In0 := WORD#16#00, In1 := WORD#16#02); END_IF;
IF P_On AND NOT MotS_CCW THEN MotS_MV := SEL(G := MotS_CW, In0 := WORD#16#00, In1 := WORD#16#01); END_IF;
IF P_On AND NOT MotS_CW THEN MotS_MV := SEL(G := MotS_CCW, In0 := WORD#16#00, In1 := WORD#16#02); END_IF;
(* Rung 15 *)
STP_SOL := Stopper_SOL[0] OR Stopper_SOL[1];

